(* IEC 61131-3 sources: deprecated-refusr-repo/samples (part 3) *)

(* ---- 2-MUX_whoso-sours-stout.st ---- *)
(*
This code implements a shuffled multiplexer with 2 control bits.
The control bits are: Data[3], Data[2]
The input bits are: Data[5], Data[1], Data[6], Data[4]

The symbolic expression is:
(((~(~(D[3]) & ~(D[2])) | D[5]) & (~(D[3] & ~(D[2])) | D[1])) & (~(~(D[3]) & D[2]) | D[6])) & (~(D[3] & D[2]) | D[4])

*)

FUNCTION_BLOCK F_CollectInput
  VAR_IN_OUT
      Data : ARRAY[1..10] OF BOOL;
  END_VAR
  VAR_INPUT
      TICK  : BOOL := 0;
      IN1   : BOOL := 0;
      IN2   : BOOL := 0;
      IN3   : BOOL := 0;
      IN4   : BOOL := 0;
      IN5   : BOOL := 0;
      RESET : BOOL := FALSE;
  END_VAR
  VAR_OUTPUT
      Finished : BOOL;
  END_VAR
  VAR
      j    : USINT := 1;
      tock : BOOL  := 0;
  END_VAR
  IF NOT RESET AND tock = NOT TICK THEN
      Data[j]   := IN1;
      Data[j+1] := IN2;
      Data[j+2] := IN3;
      Data[j+3] := IN4;
      Data[j+4] := IN5;
      j := j + 5;
      tock := TICK;
  ELSE
      j := 1;
      tock := 0;
  END_IF;
  Finished := (j > 10);
END_FUNCTION_BLOCK

PROGRAM Boiler
  VAR
    Data  : ARRAY[1..10] OF BOOL;
    Ready : BOOL;
    CollectInput : F_CollectInput;
  END_VAR
  VAR
    TICK     AT %IX1.0 : BOOL;
    IN1      AT %IX0.3 : BOOL;
    IN2      AT %IX0.4 : BOOL;
    IN3      AT %IX0.5 : BOOL;
    IN4      AT %IX0.6 : BOOL;
    IN5      AT %IX0.7 : BOOL;
    OutReady AT %QX0.0 : BOOL := FALSE;
    FeedNext AT %QX0.1 : BOOL := FALSE;
    Out      AT %QX0.2 : BOOL;
  END_VAR
  CollectInput(TICK:=TICK, IN1:=IN1, IN2:=IN2, IN3:=IN3, IN4:=IN4, IN5:=IN5);
  Ready := CollectInput.Finished;
  FeedNext := 1;
  IF Ready THEN
    Out := (((((NOT ((NOT D[3]) AND (NOT D[2]))) OR D[5]) AND ((NOT (D[3] AND (NOT D[2]))) OR D[1])) AND ((NOT ((NOT D[3]) AND D[2])) OR D[6])) AND ((NOT (D[3] AND D[2])) OR D[4]));
    OutReady := 1;
    CollectInput(RESET:=TRUE);
  END_IF;
END_PROGRAM

CONFIGURATION Config0
  RESOURCE Res0 ON PLC
    TASK task0(INTERVAL := T#20ms,PRIORITY := 0);
    PROGRAM instance0 WITH task0 : Boiler;
  END_RESOURCE
END_CONFIGURATION

(* ---- 2-MUX_wimpy-lubra-dopes.st ---- *)
(*
This code implements a shuffled multiplexer with 2 control bits.
The control bits are: Data[1], Data[5]
The input bits are: Data[3], Data[2], Data[4], Data[6]

The symbolic expression is:
(((~(~(D[1]) & ~(D[5])) | D[3]) & (~(D[1] & ~(D[5])) | D[2])) & (~(~(D[1]) & D[5]) | D[4])) & (~(D[1] & D[5]) | D[6])

*)

FUNCTION_BLOCK F_CollectInput
  VAR_IN_OUT
      Data : ARRAY[1..10] OF BOOL;
  END_VAR
  VAR_INPUT
      TICK  : BOOL := 0;
      IN1   : BOOL := 0;
      IN2   : BOOL := 0;
      IN3   : BOOL := 0;
      IN4   : BOOL := 0;
      IN5   : BOOL := 0;
      RESET : BOOL := FALSE;
  END_VAR
  VAR_OUTPUT
      Finished : BOOL;
  END_VAR
  VAR
      j    : USINT := 1;
      tock : BOOL  := 0;
  END_VAR
  IF NOT RESET AND tock = NOT TICK THEN
      Data[j]   := IN1;
      Data[j+1] := IN2;
      Data[j+2] := IN3;
      Data[j+3] := IN4;
      Data[j+4] := IN5;
      j := j + 5;
      tock := TICK;
  ELSE
      j := 1;
      tock := 0;
  END_IF;
  Finished := (j > 10);
END_FUNCTION_BLOCK

PROGRAM Boiler
  VAR
    Data  : ARRAY[1..10] OF BOOL;
    Ready : BOOL;
    CollectInput : F_CollectInput;
  END_VAR
  VAR
    TICK     AT %IX1.0 : BOOL;
    IN1      AT %IX0.3 : BOOL;
    IN2      AT %IX0.4 : BOOL;
    IN3      AT %IX0.5 : BOOL;
    IN4      AT %IX0.6 : BOOL;
    IN5      AT %IX0.7 : BOOL;
    OutReady AT %QX0.0 : BOOL := FALSE;
    FeedNext AT %QX0.1 : BOOL := FALSE;
    Out      AT %QX0.2 : BOOL;
  END_VAR
  CollectInput(TICK:=TICK, IN1:=IN1, IN2:=IN2, IN3:=IN3, IN4:=IN4, IN5:=IN5);
  Ready := CollectInput.Finished;
  FeedNext := 1;
  IF Ready THEN
    Out := (((((NOT ((NOT D[1]) AND (NOT D[5]))) OR D[3]) AND ((NOT (D[1] AND (NOT D[5]))) OR D[2])) AND ((NOT ((NOT D[1]) AND D[5])) OR D[4])) AND ((NOT (D[1] AND D[5])) OR D[6]));
    OutReady := 1;
    CollectInput(RESET:=TRUE);
  END_IF;
END_PROGRAM

CONFIGURATION Config0
  RESOURCE Res0 ON PLC
    TASK task0(INTERVAL := T#20ms,PRIORITY := 0);
    PROGRAM instance0 WITH task0 : Boiler;
  END_RESOURCE
END_CONFIGURATION

(* ---- 2-MUX_wolds-gists-resay.st ---- *)
(*
This code implements a shuffled multiplexer with 2 control bits.
The control bits are: Data[4], Data[2]
The input bits are: Data[5], Data[1], Data[3], Data[6]

The symbolic expression is:
(((~(~(D[4]) & ~(D[2])) | D[5]) & (~(D[4] & ~(D[2])) | D[1])) & (~(~(D[4]) & D[2]) | D[3])) & (~(D[4] & D[2]) | D[6])

*)

FUNCTION_BLOCK F_CollectInput
  VAR_IN_OUT
      Data : ARRAY[1..10] OF BOOL;
  END_VAR
  VAR_INPUT
      TICK  : BOOL := 0;
      IN1   : BOOL := 0;
      IN2   : BOOL := 0;
      IN3   : BOOL := 0;
      IN4   : BOOL := 0;
      IN5   : BOOL := 0;
      RESET : BOOL := FALSE;
  END_VAR
  VAR_OUTPUT
      Finished : BOOL;
  END_VAR
  VAR
      j    : USINT := 1;
      tock : BOOL  := 0;
  END_VAR
  IF NOT RESET AND tock = NOT TICK THEN
      Data[j]   := IN1;
      Data[j+1] := IN2;
      Data[j+2] := IN3;
      Data[j+3] := IN4;
      Data[j+4] := IN5;
      j := j + 5;
      tock := TICK;
  ELSE
      j := 1;
      tock := 0;
  END_IF;
  Finished := (j > 10);
END_FUNCTION_BLOCK

PROGRAM Boiler
  VAR
    Data  : ARRAY[1..10] OF BOOL;
    Ready : BOOL;
    CollectInput : F_CollectInput;
  END_VAR
  VAR
    TICK     AT %IX1.0 : BOOL;
    IN1      AT %IX0.3 : BOOL;
    IN2      AT %IX0.4 : BOOL;
    IN3      AT %IX0.5 : BOOL;
    IN4      AT %IX0.6 : BOOL;
    IN5      AT %IX0.7 : BOOL;
    OutReady AT %QX0.0 : BOOL := FALSE;
    FeedNext AT %QX0.1 : BOOL := FALSE;
    Out      AT %QX0.2 : BOOL;
  END_VAR
  CollectInput(TICK:=TICK, IN1:=IN1, IN2:=IN2, IN3:=IN3, IN4:=IN4, IN5:=IN5);
  Ready := CollectInput.Finished;
  FeedNext := 1;
  IF Ready THEN
    Out := (((((NOT ((NOT D[4]) AND (NOT D[2]))) OR D[5]) AND ((NOT (D[4] AND (NOT D[2]))) OR D[1])) AND ((NOT ((NOT D[4]) AND D[2])) OR D[3])) AND ((NOT (D[4] AND D[2])) OR D[6]));
    OutReady := 1;
    CollectInput(RESET:=TRUE);
  END_IF;
END_PROGRAM

CONFIGURATION Config0
  RESOURCE Res0 ON PLC
    TASK task0(INTERVAL := T#20ms,PRIORITY := 0);
    PROGRAM instance0 WITH task0 : Boiler;
  END_RESOURCE
END_CONFIGURATION

(* ---- 2-MUX_yella-trams-woken.st ---- *)
(*
This code implements a shuffled multiplexer with 2 control bits.
The control bits are: Data[1], Data[2]
The input bits are: Data[3], Data[5], Data[6], Data[4]

The symbolic expression is:
(((~(~(D[1]) & ~(D[2])) | D[3]) & (~(D[1] & ~(D[2])) | D[5])) & (~(~(D[1]) & D[2]) | D[6])) & (~(D[1] & D[2]) | D[4])

*)

FUNCTION_BLOCK F_CollectInput
  VAR_IN_OUT
      Data : ARRAY[1..10] OF BOOL;
  END_VAR
  VAR_INPUT
      TICK  : BOOL := 0;
      IN1   : BOOL := 0;
      IN2   : BOOL := 0;
      IN3   : BOOL := 0;
      IN4   : BOOL := 0;
      IN5   : BOOL := 0;
      RESET : BOOL := FALSE;
  END_VAR
  VAR_OUTPUT
      Finished : BOOL;
  END_VAR
  VAR
      j    : USINT := 1;
      tock : BOOL  := 0;
  END_VAR
  IF NOT RESET AND tock = NOT TICK THEN
      Data[j]   := IN1;
      Data[j+1] := IN2;
      Data[j+2] := IN3;
      Data[j+3] := IN4;
      Data[j+4] := IN5;
      j := j + 5;
      tock := TICK;
  ELSE
      j := 1;
      tock := 0;
  END_IF;
  Finished := (j > 10);
END_FUNCTION_BLOCK

PROGRAM Boiler
  VAR
    Data  : ARRAY[1..10] OF BOOL;
    Ready : BOOL;
    CollectInput : F_CollectInput;
  END_VAR
  VAR
    TICK     AT %IX1.0 : BOOL;
    IN1      AT %IX0.3 : BOOL;
    IN2      AT %IX0.4 : BOOL;
    IN3      AT %IX0.5 : BOOL;
    IN4      AT %IX0.6 : BOOL;
    IN5      AT %IX0.7 : BOOL;
    OutReady AT %QX0.0 : BOOL := FALSE;
    FeedNext AT %QX0.1 : BOOL := FALSE;
    Out      AT %QX0.2 : BOOL;
  END_VAR
  CollectInput(TICK:=TICK, IN1:=IN1, IN2:=IN2, IN3:=IN3, IN4:=IN4, IN5:=IN5);
  Ready := CollectInput.Finished;
  FeedNext := 1;
  IF Ready THEN
    Out := (((((NOT ((NOT D[1]) AND (NOT D[2]))) OR D[3]) AND ((NOT (D[1] AND (NOT D[2]))) OR D[5])) AND ((NOT ((NOT D[1]) AND D[2])) OR D[6])) AND ((NOT (D[1] AND D[2])) OR D[4]));
    OutReady := 1;
    CollectInput(RESET:=TRUE);
  END_IF;
END_PROGRAM

CONFIGURATION Config0
  RESOURCE Res0 ON PLC
    TASK task0(INTERVAL := T#20ms,PRIORITY := 0);
    PROGRAM instance0 WITH task0 : Boiler;
  END_RESOURCE
END_CONFIGURATION

(* ---- 2-MUX_yoyos-blast-cameo.st ---- *)
(*
This code implements a shuffled multiplexer with 2 control bits.
The control bits are: Data[3], Data[2]
The input bits are: Data[1], Data[4], Data[5], Data[6]

The symbolic expression is:
(((~(~(D[3]) & ~(D[2])) | D[1]) & (~(D[3] & ~(D[2])) | D[4])) & (~(~(D[3]) & D[2]) | D[5])) & (~(D[3] & D[2]) | D[6])

*)

FUNCTION_BLOCK F_CollectInput
  VAR_IN_OUT
      Data : ARRAY[1..10] OF BOOL;
  END_VAR
  VAR_INPUT
      TICK  : BOOL := 0;
      IN1   : BOOL := 0;
      IN2   : BOOL := 0;
      IN3   : BOOL := 0;
      IN4   : BOOL := 0;
      IN5   : BOOL := 0;
      RESET : BOOL := FALSE;
  END_VAR
  VAR_OUTPUT
      Finished : BOOL;
  END_VAR
  VAR
      j    : USINT := 1;
      tock : BOOL  := 0;
  END_VAR
  IF NOT RESET AND tock = NOT TICK THEN
      Data[j]   := IN1;
      Data[j+1] := IN2;
      Data[j+2] := IN3;
      Data[j+3] := IN4;
      Data[j+4] := IN5;
      j := j + 5;
      tock := TICK;
  ELSE
      j := 1;
      tock := 0;
  END_IF;
  Finished := (j > 10);
END_FUNCTION_BLOCK

PROGRAM Boiler
  VAR
    Data  : ARRAY[1..10] OF BOOL;
    Ready : BOOL;
    CollectInput : F_CollectInput;
  END_VAR
  VAR
    TICK     AT %IX1.0 : BOOL;
    IN1      AT %IX0.3 : BOOL;
    IN2      AT %IX0.4 : BOOL;
    IN3      AT %IX0.5 : BOOL;
    IN4      AT %IX0.6 : BOOL;
    IN5      AT %IX0.7 : BOOL;
    OutReady AT %QX0.0 : BOOL := FALSE;
    FeedNext AT %QX0.1 : BOOL := FALSE;
    Out      AT %QX0.2 : BOOL;
  END_VAR
  CollectInput(TICK:=TICK, IN1:=IN1, IN2:=IN2, IN3:=IN3, IN4:=IN4, IN5:=IN5);
  Ready := CollectInput.Finished;
  FeedNext := 1;
  IF Ready THEN
    Out := (((((NOT ((NOT D[3]) AND (NOT D[2]))) OR D[1]) AND ((NOT (D[3] AND (NOT D[2]))) OR D[4])) AND ((NOT ((NOT D[3]) AND D[2])) OR D[5])) AND ((NOT (D[3] AND D[2])) OR D[6]));
    OutReady := 1;
    CollectInput(RESET:=TRUE);
  END_IF;
END_PROGRAM

CONFIGURATION Config0
  RESOURCE Res0 ON PLC
    TASK task0(INTERVAL := T#20ms,PRIORITY := 0);
    PROGRAM instance0 WITH task0 : Boiler;
  END_RESOURCE
END_CONFIGURATION

(* ---- 2-MUX_yurts-tippy-sayer.st ---- *)
(*
This code implements a shuffled multiplexer with 2 control bits.
The control bits are: Data[3], Data[1]
The input bits are: Data[4], Data[2], Data[5], Data[6]

The symbolic expression is:
(((~(~(D[3]) & ~(D[1])) | D[4]) & (~(D[3] & ~(D[1])) | D[2])) & (~(~(D[3]) & D[1]) | D[5])) & (~(D[3] & D[1]) | D[6])

*)

FUNCTION_BLOCK F_CollectInput
  VAR_IN_OUT
      Data : ARRAY[1..10] OF BOOL;
  END_VAR
  VAR_INPUT
      TICK  : BOOL := 0;
      IN1   : BOOL := 0;
      IN2   : BOOL := 0;
      IN3   : BOOL := 0;
      IN4   : BOOL := 0;
      IN5   : BOOL := 0;
      RESET : BOOL := FALSE;
  END_VAR
  VAR_OUTPUT
      Finished : BOOL;
  END_VAR
  VAR
      j    : USINT := 1;
      tock : BOOL  := 0;
  END_VAR
  IF NOT RESET AND tock = NOT TICK THEN
      Data[j]   := IN1;
      Data[j+1] := IN2;
      Data[j+2] := IN3;
      Data[j+3] := IN4;
      Data[j+4] := IN5;
      j := j + 5;
      tock := TICK;
  ELSE
      j := 1;
      tock := 0;
  END_IF;
  Finished := (j > 10);
END_FUNCTION_BLOCK

PROGRAM Boiler
  VAR
    Data  : ARRAY[1..10] OF BOOL;
    Ready : BOOL;
    CollectInput : F_CollectInput;
  END_VAR
  VAR
    TICK     AT %IX1.0 : BOOL;
    IN1      AT %IX0.3 : BOOL;
    IN2      AT %IX0.4 : BOOL;
    IN3      AT %IX0.5 : BOOL;
    IN4      AT %IX0.6 : BOOL;
    IN5      AT %IX0.7 : BOOL;
    OutReady AT %QX0.0 : BOOL := FALSE;
    FeedNext AT %QX0.1 : BOOL := FALSE;
    Out      AT %QX0.2 : BOOL;
  END_VAR
  CollectInput(TICK:=TICK, IN1:=IN1, IN2:=IN2, IN3:=IN3, IN4:=IN4, IN5:=IN5);
  Ready := CollectInput.Finished;
  FeedNext := 1;
  IF Ready THEN
    Out := (((((NOT ((NOT D[3]) AND (NOT D[1]))) OR D[4]) AND ((NOT (D[3] AND (NOT D[1]))) OR D[2])) AND ((NOT ((NOT D[3]) AND D[1])) OR D[5])) AND ((NOT (D[3] AND D[1])) OR D[6]));
    OutReady := 1;
    CollectInput(RESET:=TRUE);
  END_IF;
END_PROGRAM

CONFIGURATION Config0
  RESOURCE Res0 ON PLC
    TASK task0(INTERVAL := T#20ms,PRIORITY := 0);
    PROGRAM instance0 WITH task0 : Boiler;
  END_RESOURCE
END_CONFIGURATION

(* ---- 2-MUX_zebus-trove-teals.st ---- *)
(*
This code implements a shuffled multiplexer with 2 control bits.
The control bits are: Data[2], Data[1]
The input bits are: Data[5], Data[6], Data[3], Data[4]

The symbolic expression is:
(((~(~(D[2]) & ~(D[1])) | D[5]) & (~(D[2] & ~(D[1])) | D[6])) & (~(~(D[2]) & D[1]) | D[3])) & (~(D[2] & D[1]) | D[4])

*)

FUNCTION_BLOCK F_CollectInput
  VAR_IN_OUT
      Data : ARRAY[1..10] OF BOOL;
  END_VAR
  VAR_INPUT
      TICK  : BOOL := 0;
      IN1   : BOOL := 0;
      IN2   : BOOL := 0;
      IN3   : BOOL := 0;
      IN4   : BOOL := 0;
      IN5   : BOOL := 0;
      RESET : BOOL := FALSE;
  END_VAR
  VAR_OUTPUT
      Finished : BOOL;
  END_VAR
  VAR
      j    : USINT := 1;
      tock : BOOL  := 0;
  END_VAR
  IF NOT RESET AND tock = NOT TICK THEN
      Data[j]   := IN1;
      Data[j+1] := IN2;
      Data[j+2] := IN3;
      Data[j+3] := IN4;
      Data[j+4] := IN5;
      j := j + 5;
      tock := TICK;
  ELSE
      j := 1;
      tock := 0;
  END_IF;
  Finished := (j > 10);
END_FUNCTION_BLOCK

PROGRAM Boiler
  VAR
    Data  : ARRAY[1..10] OF BOOL;
    Ready : BOOL;
    CollectInput : F_CollectInput;
  END_VAR
  VAR
    TICK     AT %IX1.0 : BOOL;
    IN1      AT %IX0.3 : BOOL;
    IN2      AT %IX0.4 : BOOL;
    IN3      AT %IX0.5 : BOOL;
    IN4      AT %IX0.6 : BOOL;
    IN5      AT %IX0.7 : BOOL;
    OutReady AT %QX0.0 : BOOL := FALSE;
    FeedNext AT %QX0.1 : BOOL := FALSE;
    Out      AT %QX0.2 : BOOL;
  END_VAR
  CollectInput(TICK:=TICK, IN1:=IN1, IN2:=IN2, IN3:=IN3, IN4:=IN4, IN5:=IN5);
  Ready := CollectInput.Finished;
  FeedNext := 1;
  IF Ready THEN
    Out := (((((NOT ((NOT D[2]) AND (NOT D[1]))) OR D[5]) AND ((NOT (D[2] AND (NOT D[1]))) OR D[6])) AND ((NOT ((NOT D[2]) AND D[1])) OR D[3])) AND ((NOT (D[2] AND D[1])) OR D[4]));
    OutReady := 1;
    CollectInput(RESET:=TRUE);
  END_IF;
END_PROGRAM

CONFIGURATION Config0
  RESOURCE Res0 ON PLC
    TASK task0(INTERVAL := T#20ms,PRIORITY := 0);
    PROGRAM instance0 WITH task0 : Boiler;
  END_RESOURCE
END_CONFIGURATION

(* ---- 2-MUX_zebus-whiny-fares.st ---- *)
(*
This code implements a shuffled multiplexer with 2 control bits.
The control bits are: Data[1], Data[2]
The input bits are: Data[3], Data[4], Data[5], Data[6]

The symbolic expression is:
(((~(~(D[1]) & ~(D[2])) | D[3]) & (~(D[1] & ~(D[2])) | D[4])) & (~(~(D[1]) & D[2]) | D[5])) & (~(D[1] & D[2]) | D[6])

*)

FUNCTION_BLOCK F_CollectInput
  VAR_IN_OUT
      Data : ARRAY[1..10] OF BOOL;
  END_VAR
  VAR_INPUT
      TICK  : BOOL := 0;
      IN1   : BOOL := 0;
      IN2   : BOOL := 0;
      IN3   : BOOL := 0;
      IN4   : BOOL := 0;
      IN5   : BOOL := 0;
      RESET : BOOL := FALSE;
  END_VAR
  VAR_OUTPUT
      Finished : BOOL;
  END_VAR
  VAR
      j    : USINT := 1;
      tock : BOOL  := 0;
  END_VAR
  IF NOT RESET AND tock = NOT TICK THEN
      Data[j]   := IN1;
      Data[j+1] := IN2;
      Data[j+2] := IN3;
      Data[j+3] := IN4;
      Data[j+4] := IN5;
      j := j + 5;
      tock := TICK;
  ELSE
      j := 1;
      tock := 0;
  END_IF;
  Finished := (j > 10);
END_FUNCTION_BLOCK

PROGRAM Boiler
  VAR
    Data  : ARRAY[1..10] OF BOOL;
    Ready : BOOL;
    CollectInput : F_CollectInput;
  END_VAR
  VAR
    TICK     AT %IX1.0 : BOOL;
    IN1      AT %IX0.3 : BOOL;
    IN2      AT %IX0.4 : BOOL;
    IN3      AT %IX0.5 : BOOL;
    IN4      AT %IX0.6 : BOOL;
    IN5      AT %IX0.7 : BOOL;
    OutReady AT %QX0.0 : BOOL := FALSE;
    FeedNext AT %QX0.1 : BOOL := FALSE;
    Out      AT %QX0.2 : BOOL;
  END_VAR
  CollectInput(TICK:=TICK, IN1:=IN1, IN2:=IN2, IN3:=IN3, IN4:=IN4, IN5:=IN5);
  Ready := CollectInput.Finished;
  FeedNext := 1;
  IF Ready THEN
    Out := (((((NOT ((NOT D[1]) AND (NOT D[2]))) OR D[3]) AND ((NOT (D[1] AND (NOT D[2]))) OR D[4])) AND ((NOT ((NOT D[1]) AND D[2])) OR D[5])) AND ((NOT (D[1] AND D[2])) OR D[6]));
    OutReady := 1;
    CollectInput(RESET:=TRUE);
  END_IF;
END_PROGRAM

CONFIGURATION Config0
  RESOURCE Res0 ON PLC
    TASK task0(INTERVAL := T#20ms,PRIORITY := 0);
    PROGRAM instance0 WITH task0 : Boiler;
  END_RESOURCE
END_CONFIGURATION

(* ---- 3-MUX_acked-palls-seven.st ---- *)
(*
This code implements a shuffled multiplexer with 3 control bits.
The control bits are: Data[2], Data[1], Data[3]
The input bits are: Data[4], Data[6], Data[7], Data[5], Data[8], Data[9], Data[11], Data[10]

The symbolic expression is:
(((((((~((~(D[2]) & ~(D[1])) & ~(D[3])) | D[4]) & (~((D[2] & ~(D[1])) & ~(D[3])) | D[6])) & (~((~(D[2]) & D[1]) & ~(D[3])) | D[7])) & (~((D[2] & D[1]) & ~(D[3])) | D[5])) & (~((~(D[2]) & ~(D[1])) & D[3]) | D[8])) & (~((D[2] & ~(D[1])) & D[3]) | D[9])) & (~((~(D[2]) & D[1]) & D[3]) | D[11])) & (~((D[2] & D[1]) & D[3]) | D[10])

*)

FUNCTION_BLOCK F_CollectInput
  VAR_IN_OUT
      Data : ARRAY[1..15] OF BOOL;
  END_VAR
  VAR_INPUT
      TICK  : BOOL := 0;
      IN1   : BOOL := 0;
      IN2   : BOOL := 0;
      IN3   : BOOL := 0;
      IN4   : BOOL := 0;
      IN5   : BOOL := 0;
      RESET : BOOL := FALSE;
  END_VAR
  VAR_OUTPUT
      Finished : BOOL;
  END_VAR
  VAR
      j    : USINT := 1;
      tock : BOOL  := 0;
  END_VAR
  IF NOT RESET AND tock = NOT TICK THEN
      Data[j]   := IN1;
      Data[j+1] := IN2;
      Data[j+2] := IN3;
      Data[j+3] := IN4;
      Data[j+4] := IN5;
      j := j + 5;
      tock := TICK;
  ELSE
      j := 1;
      tock := 0;
  END_IF;
  Finished := (j > 15);
END_FUNCTION_BLOCK

PROGRAM Boiler
  VAR
    Data  : ARRAY[1..15] OF BOOL;
    Ready : BOOL;
    CollectInput : F_CollectInput;
  END_VAR
  VAR
    TICK     AT %IX1.0 : BOOL;
    IN1      AT %IX0.3 : BOOL;
    IN2      AT %IX0.4 : BOOL;
    IN3      AT %IX0.5 : BOOL;
    IN4      AT %IX0.6 : BOOL;
    IN5      AT %IX0.7 : BOOL;
    OutReady AT %QX0.0 : BOOL := FALSE;
    FeedNext AT %QX0.1 : BOOL := FALSE;
    Out      AT %QX0.2 : BOOL;
  END_VAR
  CollectInput(TICK:=TICK, IN1:=IN1, IN2:=IN2, IN3:=IN3, IN4:=IN4, IN5:=IN5);
  Ready := CollectInput.Finished;
  FeedNext := 1;
  IF Ready THEN
    Out := (((((((((NOT (((NOT D[2]) AND (NOT D[1])) AND (NOT D[3]))) OR D[4]) AND ((NOT ((D[2] AND (NOT D[1])) AND (NOT D[3]))) OR D[6])) AND ((NOT (((NOT D[2]) AND D[1]) AND (NOT D[3]))) OR D[7])) AND ((NOT ((D[2] AND D[1]) AND (NOT D[3]))) OR D[5])) AND ((NOT (((NOT D[2]) AND (NOT D[1])) AND D[3])) OR D[8])) AND ((NOT ((D[2] AND (NOT D[1])) AND D[3])) OR D[9])) AND ((NOT (((NOT D[2]) AND D[1]) AND D[3])) OR D[11])) AND ((NOT ((D[2] AND D[1]) AND D[3])) OR D[10]));
    OutReady := 1;
    CollectInput(RESET:=TRUE);
  END_IF;
END_PROGRAM

CONFIGURATION Config0
  RESOURCE Res0 ON PLC
    TASK task0(INTERVAL := T#20ms,PRIORITY := 0);
    PROGRAM instance0 WITH task0 : Boiler;
  END_RESOURCE
END_CONFIGURATION

(* ---- 3-MUX_alums-tends-demon.st ---- *)
(*
This code implements a shuffled multiplexer with 3 control bits.
The control bits are: Data[1], Data[3], Data[6]
The input bits are: Data[4], Data[9], Data[5], Data[2], Data[7], Data[8], Data[10], Data[11]

The symbolic expression is:
(((((((~((~(D[1]) & ~(D[3])) & ~(D[6])) | D[4]) & (~((D[1] & ~(D[3])) & ~(D[6])) | D[9])) & (~((~(D[1]) & D[3]) & ~(D[6])) | D[5])) & (~((D[1] & D[3]) & ~(D[6])) | D[2])) & (~((~(D[1]) & ~(D[3])) & D[6]) | D[7])) & (~((D[1] & ~(D[3])) & D[6]) | D[8])) & (~((~(D[1]) & D[3]) & D[6]) | D[10])) & (~((D[1] & D[3]) & D[6]) | D[11])

*)

FUNCTION_BLOCK F_CollectInput
  VAR_IN_OUT
      Data : ARRAY[1..15] OF BOOL;
  END_VAR
  VAR_INPUT
      TICK  : BOOL := 0;
      IN1   : BOOL := 0;
      IN2   : BOOL := 0;
      IN3   : BOOL := 0;
      IN4   : BOOL := 0;
      IN5   : BOOL := 0;
      RESET : BOOL := FALSE;
  END_VAR
  VAR_OUTPUT
      Finished : BOOL;
  END_VAR
  VAR
      j    : USINT := 1;
      tock : BOOL  := 0;
  END_VAR
  IF NOT RESET AND tock = NOT TICK THEN
      Data[j]   := IN1;
      Data[j+1] := IN2;
      Data[j+2] := IN3;
      Data[j+3] := IN4;
      Data[j+4] := IN5;
      j := j + 5;
      tock := TICK;
  ELSE
      j := 1;
      tock := 0;
  END_IF;
  Finished := (j > 15);
END_FUNCTION_BLOCK

PROGRAM Boiler
  VAR
    Data  : ARRAY[1..15] OF BOOL;
    Ready : BOOL;
    CollectInput : F_CollectInput;
  END_VAR
  VAR
    TICK     AT %IX1.0 : BOOL;
    IN1      AT %IX0.3 : BOOL;
    IN2      AT %IX0.4 : BOOL;
    IN3      AT %IX0.5 : BOOL;
    IN4      AT %IX0.6 : BOOL;
    IN5      AT %IX0.7 : BOOL;
    OutReady AT %QX0.0 : BOOL := FALSE;
    FeedNext AT %QX0.1 : BOOL := FALSE;
    Out      AT %QX0.2 : BOOL;
  END_VAR
  CollectInput(TICK:=TICK, IN1:=IN1, IN2:=IN2, IN3:=IN3, IN4:=IN4, IN5:=IN5);
  Ready := CollectInput.Finished;
  FeedNext := 1;
  IF Ready THEN
    Out := (((((((((NOT (((NOT D[1]) AND (NOT D[3])) AND (NOT D[6]))) OR D[4]) AND ((NOT ((D[1] AND (NOT D[3])) AND (NOT D[6]))) OR D[9])) AND ((NOT (((NOT D[1]) AND D[3]) AND (NOT D[6]))) OR D[5])) AND ((NOT ((D[1] AND D[3]) AND (NOT D[6]))) OR D[2])) AND ((NOT (((NOT D[1]) AND (NOT D[3])) AND D[6])) OR D[7])) AND ((NOT ((D[1] AND (NOT D[3])) AND D[6])) OR D[8])) AND ((NOT (((NOT D[1]) AND D[3]) AND D[6])) OR D[10])) AND ((NOT ((D[1] AND D[3]) AND D[6])) OR D[11]));
    OutReady := 1;
    CollectInput(RESET:=TRUE);
  END_IF;
END_PROGRAM

CONFIGURATION Config0
  RESOURCE Res0 ON PLC
    TASK task0(INTERVAL := T#20ms,PRIORITY := 0);
    PROGRAM instance0 WITH task0 : Boiler;
  END_RESOURCE
END_CONFIGURATION

(* ---- 3-MUX_annex-saucy-first.st ---- *)
(*
This code implements a shuffled multiplexer with 3 control bits.
The control bits are: Data[2], Data[1], Data[5]
The input bits are: Data[3], Data[6], Data[4], Data[7], Data[8], Data[9], Data[10], Data[11]

The symbolic expression is:
(((((((~((~(D[2]) & ~(D[1])) & ~(D[5])) | D[3]) & (~((D[2] & ~(D[1])) & ~(D[5])) | D[6])) & (~((~(D[2]) & D[1]) & ~(D[5])) | D[4])) & (~((D[2] & D[1]) & ~(D[5])) | D[7])) & (~((~(D[2]) & ~(D[1])) & D[5]) | D[8])) & (~((D[2] & ~(D[1])) & D[5]) | D[9])) & (~((~(D[2]) & D[1]) & D[5]) | D[10])) & (~((D[2] & D[1]) & D[5]) | D[11])

*)

FUNCTION_BLOCK F_CollectInput
  VAR_IN_OUT
      Data : ARRAY[1..15] OF BOOL;
  END_VAR
  VAR_INPUT
      TICK  : BOOL := 0;
      IN1   : BOOL := 0;
      IN2   : BOOL := 0;
      IN3   : BOOL := 0;
      IN4   : BOOL := 0;
      IN5   : BOOL := 0;
      RESET : BOOL := FALSE;
  END_VAR
  VAR_OUTPUT
      Finished : BOOL;
  END_VAR
  VAR
      j    : USINT := 1;
      tock : BOOL  := 0;
  END_VAR
  IF NOT RESET AND tock = NOT TICK THEN
      Data[j]   := IN1;
      Data[j+1] := IN2;
      Data[j+2] := IN3;
      Data[j+3] := IN4;
      Data[j+4] := IN5;
      j := j + 5;
      tock := TICK;
  ELSE
      j := 1;
      tock := 0;
  END_IF;
  Finished := (j > 15);
END_FUNCTION_BLOCK

PROGRAM Boiler
  VAR
    Data  : ARRAY[1..15] OF BOOL;
    Ready : BOOL;
    CollectInput : F_CollectInput;
  END_VAR
  VAR
    TICK     AT %IX1.0 : BOOL;
    IN1      AT %IX0.3 : BOOL;
    IN2      AT %IX0.4 : BOOL;
    IN3      AT %IX0.5 : BOOL;
    IN4      AT %IX0.6 : BOOL;
    IN5      AT %IX0.7 : BOOL;
    OutReady AT %QX0.0 : BOOL := FALSE;
    FeedNext AT %QX0.1 : BOOL := FALSE;
    Out      AT %QX0.2 : BOOL;
  END_VAR
  CollectInput(TICK:=TICK, IN1:=IN1, IN2:=IN2, IN3:=IN3, IN4:=IN4, IN5:=IN5);
  Ready := CollectInput.Finished;
  FeedNext := 1;
  IF Ready THEN
    Out := (((((((((NOT (((NOT D[2]) AND (NOT D[1])) AND (NOT D[5]))) OR D[3]) AND ((NOT ((D[2] AND (NOT D[1])) AND (NOT D[5]))) OR D[6])) AND ((NOT (((NOT D[2]) AND D[1]) AND (NOT D[5]))) OR D[4])) AND ((NOT ((D[2] AND D[1]) AND (NOT D[5]))) OR D[7])) AND ((NOT (((NOT D[2]) AND (NOT D[1])) AND D[5])) OR D[8])) AND ((NOT ((D[2] AND (NOT D[1])) AND D[5])) OR D[9])) AND ((NOT (((NOT D[2]) AND D[1]) AND D[5])) OR D[10])) AND ((NOT ((D[2] AND D[1]) AND D[5])) OR D[11]));
    OutReady := 1;
    CollectInput(RESET:=TRUE);
  END_IF;
END_PROGRAM

CONFIGURATION Config0
  RESOURCE Res0 ON PLC
    TASK task0(INTERVAL := T#20ms,PRIORITY := 0);
    PROGRAM instance0 WITH task0 : Boiler;
  END_RESOURCE
END_CONFIGURATION

(* ---- 3-MUX_antic-lucks-mould.st ---- *)
(*
This code implements a shuffled multiplexer with 3 control bits.
The control bits are: Data[2], Data[7], Data[1]
The input bits are: Data[3], Data[5], Data[6], Data[4], Data[8], Data[9], Data[10], Data[11]

The symbolic expression is:
(((((((~((~(D[2]) & ~(D[7])) & ~(D[1])) | D[3]) & (~((D[2] & ~(D[7])) & ~(D[1])) | D[5])) & (~((~(D[2]) & D[7]) & ~(D[1])) | D[6])) & (~((D[2] & D[7]) & ~(D[1])) | D[4])) & (~((~(D[2]) & ~(D[7])) & D[1]) | D[8])) & (~((D[2] & ~(D[7])) & D[1]) | D[9])) & (~((~(D[2]) & D[7]) & D[1]) | D[10])) & (~((D[2] & D[7]) & D[1]) | D[11])

*)

FUNCTION_BLOCK F_CollectInput
  VAR_IN_OUT
      Data : ARRAY[1..15] OF BOOL;
  END_VAR
  VAR_INPUT
      TICK  : BOOL := 0;
      IN1   : BOOL := 0;
      IN2   : BOOL := 0;
      IN3   : BOOL := 0;
      IN4   : BOOL := 0;
      IN5   : BOOL := 0;
      RESET : BOOL := FALSE;
  END_VAR
  VAR_OUTPUT
      Finished : BOOL;
  END_VAR
  VAR
      j    : USINT := 1;
      tock : BOOL  := 0;
  END_VAR
  IF NOT RESET AND tock = NOT TICK THEN
      Data[j]   := IN1;
      Data[j+1] := IN2;
      Data[j+2] := IN3;
      Data[j+3] := IN4;
      Data[j+4] := IN5;
      j := j + 5;
      tock := TICK;
  ELSE
      j := 1;
      tock := 0;
  END_IF;
  Finished := (j > 15);
END_FUNCTION_BLOCK

PROGRAM Boiler
  VAR
    Data  : ARRAY[1..15] OF BOOL;
    Ready : BOOL;
    CollectInput : F_CollectInput;
  END_VAR
  VAR
    TICK     AT %IX1.0 : BOOL;
    IN1      AT %IX0.3 : BOOL;
    IN2      AT %IX0.4 : BOOL;
    IN3      AT %IX0.5 : BOOL;
    IN4      AT %IX0.6 : BOOL;
    IN5      AT %IX0.7 : BOOL;
    OutReady AT %QX0.0 : BOOL := FALSE;
    FeedNext AT %QX0.1 : BOOL := FALSE;
    Out      AT %QX0.2 : BOOL;
  END_VAR
  CollectInput(TICK:=TICK, IN1:=IN1, IN2:=IN2, IN3:=IN3, IN4:=IN4, IN5:=IN5);
  Ready := CollectInput.Finished;
  FeedNext := 1;
  IF Ready THEN
    Out := (((((((((NOT (((NOT D[2]) AND (NOT D[7])) AND (NOT D[1]))) OR D[3]) AND ((NOT ((D[2] AND (NOT D[7])) AND (NOT D[1]))) OR D[5])) AND ((NOT (((NOT D[2]) AND D[7]) AND (NOT D[1]))) OR D[6])) AND ((NOT ((D[2] AND D[7]) AND (NOT D[1]))) OR D[4])) AND ((NOT (((NOT D[2]) AND (NOT D[7])) AND D[1])) OR D[8])) AND ((NOT ((D[2] AND (NOT D[7])) AND D[1])) OR D[9])) AND ((NOT (((NOT D[2]) AND D[7]) AND D[1])) OR D[10])) AND ((NOT ((D[2] AND D[7]) AND D[1])) OR D[11]));
    OutReady := 1;
    CollectInput(RESET:=TRUE);
  END_IF;
END_PROGRAM

CONFIGURATION Config0
  RESOURCE Res0 ON PLC
    TASK task0(INTERVAL := T#20ms,PRIORITY := 0);
    PROGRAM instance0 WITH task0 : Boiler;
  END_RESOURCE
END_CONFIGURATION

(* ---- 3-MUX_apian-braes-rolls.st ---- *)
(*
This code implements a shuffled multiplexer with 3 control bits.
The control bits are: Data[2], Data[3], Data[1]
The input bits are: Data[4], Data[6], Data[5], Data[7], Data[10], Data[8], Data[9], Data[11]

The symbolic expression is:
(((((((~((~(D[2]) & ~(D[3])) & ~(D[1])) | D[4]) & (~((D[2] & ~(D[3])) & ~(D[1])) | D[6])) & (~((~(D[2]) & D[3]) & ~(D[1])) | D[5])) & (~((D[2] & D[3]) & ~(D[1])) | D[7])) & (~((~(D[2]) & ~(D[3])) & D[1]) | D[10])) & (~((D[2] & ~(D[3])) & D[1]) | D[8])) & (~((~(D[2]) & D[3]) & D[1]) | D[9])) & (~((D[2] & D[3]) & D[1]) | D[11])

*)

FUNCTION_BLOCK F_CollectInput
  VAR_IN_OUT
      Data : ARRAY[1..15] OF BOOL;
  END_VAR
  VAR_INPUT
      TICK  : BOOL := 0;
      IN1   : BOOL := 0;
      IN2   : BOOL := 0;
      IN3   : BOOL := 0;
      IN4   : BOOL := 0;
      IN5   : BOOL := 0;
      RESET : BOOL := FALSE;
  END_VAR
  VAR_OUTPUT
      Finished : BOOL;
  END_VAR
  VAR
      j    : USINT := 1;
      tock : BOOL  := 0;
  END_VAR
  IF NOT RESET AND tock = NOT TICK THEN
      Data[j]   := IN1;
      Data[j+1] := IN2;
      Data[j+2] := IN3;
      Data[j+3] := IN4;
      Data[j+4] := IN5;
      j := j + 5;
      tock := TICK;
  ELSE
      j := 1;
      tock := 0;
  END_IF;
  Finished := (j > 15);
END_FUNCTION_BLOCK

PROGRAM Boiler
  VAR
    Data  : ARRAY[1..15] OF BOOL;
    Ready : BOOL;
    CollectInput : F_CollectInput;
  END_VAR
  VAR
    TICK     AT %IX1.0 : BOOL;
    IN1      AT %IX0.3 : BOOL;
    IN2      AT %IX0.4 : BOOL;
    IN3      AT %IX0.5 : BOOL;
    IN4      AT %IX0.6 : BOOL;
    IN5      AT %IX0.7 : BOOL;
    OutReady AT %QX0.0 : BOOL := FALSE;
    FeedNext AT %QX0.1 : BOOL := FALSE;
    Out      AT %QX0.2 : BOOL;
  END_VAR
  CollectInput(TICK:=TICK, IN1:=IN1, IN2:=IN2, IN3:=IN3, IN4:=IN4, IN5:=IN5);
  Ready := CollectInput.Finished;
  FeedNext := 1;
  IF Ready THEN
    Out := (((((((((NOT (((NOT D[2]) AND (NOT D[3])) AND (NOT D[1]))) OR D[4]) AND ((NOT ((D[2] AND (NOT D[3])) AND (NOT D[1]))) OR D[6])) AND ((NOT (((NOT D[2]) AND D[3]) AND (NOT D[1]))) OR D[5])) AND ((NOT ((D[2] AND D[3]) AND (NOT D[1]))) OR D[7])) AND ((NOT (((NOT D[2]) AND (NOT D[3])) AND D[1])) OR D[10])) AND ((NOT ((D[2] AND (NOT D[3])) AND D[1])) OR D[8])) AND ((NOT (((NOT D[2]) AND D[3]) AND D[1])) OR D[9])) AND ((NOT ((D[2] AND D[3]) AND D[1])) OR D[11]));
    OutReady := 1;
    CollectInput(RESET:=TRUE);
  END_IF;
END_PROGRAM

CONFIGURATION Config0
  RESOURCE Res0 ON PLC
    TASK task0(INTERVAL := T#20ms,PRIORITY := 0);
    PROGRAM instance0 WITH task0 : Boiler;
  END_RESOURCE
END_CONFIGURATION

(* ---- 3-MUX_aping-spark-squad.st ---- *)
(*
This code implements a shuffled multiplexer with 3 control bits.
The control bits are: Data[5], Data[2], Data[1]
The input bits are: Data[4], Data[3], Data[6], Data[7], Data[8], Data[10], Data[9], Data[11]

The symbolic expression is:
(((((((~((~(D[5]) & ~(D[2])) & ~(D[1])) | D[4]) & (~((D[5] & ~(D[2])) & ~(D[1])) | D[3])) & (~((~(D[5]) & D[2]) & ~(D[1])) | D[6])) & (~((D[5] & D[2]) & ~(D[1])) | D[7])) & (~((~(D[5]) & ~(D[2])) & D[1]) | D[8])) & (~((D[5] & ~(D[2])) & D[1]) | D[10])) & (~((~(D[5]) & D[2]) & D[1]) | D[9])) & (~((D[5] & D[2]) & D[1]) | D[11])

*)

FUNCTION_BLOCK F_CollectInput
  VAR_IN_OUT
      Data : ARRAY[1..15] OF BOOL;
  END_VAR
  VAR_INPUT
      TICK  : BOOL := 0;
      IN1   : BOOL := 0;
      IN2   : BOOL := 0;
      IN3   : BOOL := 0;
      IN4   : BOOL := 0;
      IN5   : BOOL := 0;
      RESET : BOOL := FALSE;
  END_VAR
  VAR_OUTPUT
      Finished : BOOL;
  END_VAR
  VAR
      j    : USINT := 1;
      tock : BOOL  := 0;
  END_VAR
  IF NOT RESET AND tock = NOT TICK THEN
      Data[j]   := IN1;
      Data[j+1] := IN2;
      Data[j+2] := IN3;
      Data[j+3] := IN4;
      Data[j+4] := IN5;
      j := j + 5;
      tock := TICK;
  ELSE
      j := 1;
      tock := 0;
  END_IF;
  Finished := (j > 15);
END_FUNCTION_BLOCK

PROGRAM Boiler
  VAR
    Data  : ARRAY[1..15] OF BOOL;
    Ready : BOOL;
    CollectInput : F_CollectInput;
  END_VAR
  VAR
    TICK     AT %IX1.0 : BOOL;
    IN1      AT %IX0.3 : BOOL;
    IN2      AT %IX0.4 : BOOL;
    IN3      AT %IX0.5 : BOOL;
    IN4      AT %IX0.6 : BOOL;
    IN5      AT %IX0.7 : BOOL;
    OutReady AT %QX0.0 : BOOL := FALSE;
    FeedNext AT %QX0.1 : BOOL := FALSE;
    Out      AT %QX0.2 : BOOL;
  END_VAR
  CollectInput(TICK:=TICK, IN1:=IN1, IN2:=IN2, IN3:=IN3, IN4:=IN4, IN5:=IN5);
  Ready := CollectInput.Finished;
  FeedNext := 1;
  IF Ready THEN
    Out := (((((((((NOT (((NOT D[5]) AND (NOT D[2])) AND (NOT D[1]))) OR D[4]) AND ((NOT ((D[5] AND (NOT D[2])) AND (NOT D[1]))) OR D[3])) AND ((NOT (((NOT D[5]) AND D[2]) AND (NOT D[1]))) OR D[6])) AND ((NOT ((D[5] AND D[2]) AND (NOT D[1]))) OR D[7])) AND ((NOT (((NOT D[5]) AND (NOT D[2])) AND D[1])) OR D[8])) AND ((NOT ((D[5] AND (NOT D[2])) AND D[1])) OR D[10])) AND ((NOT (((NOT D[5]) AND D[2]) AND D[1])) OR D[9])) AND ((NOT ((D[5] AND D[2]) AND D[1])) OR D[11]));
    OutReady := 1;
    CollectInput(RESET:=TRUE);
  END_IF;
END_PROGRAM

CONFIGURATION Config0
  RESOURCE Res0 ON PLC
    TASK task0(INTERVAL := T#20ms,PRIORITY := 0);
    PROGRAM instance0 WITH task0 : Boiler;
  END_RESOURCE
END_CONFIGURATION

(* ---- 3-MUX_augur-aleph-tiers.st ---- *)
(*
This code implements a shuffled multiplexer with 3 control bits.
The control bits are: Data[1], Data[2], Data[10]
The input bits are: Data[4], Data[5], Data[3], Data[8], Data[6], Data[7], Data[11], Data[9]

The symbolic expression is:
(((((((~((~(D[1]) & ~(D[2])) & ~(D[10])) | D[4]) & (~((D[1] & ~(D[2])) & ~(D[10])) | D[5])) & (~((~(D[1]) & D[2]) & ~(D[10])) | D[3])) & (~((D[1] & D[2]) & ~(D[10])) | D[8])) & (~((~(D[1]) & ~(D[2])) & D[10]) | D[6])) & (~((D[1] & ~(D[2])) & D[10]) | D[7])) & (~((~(D[1]) & D[2]) & D[10]) | D[11])) & (~((D[1] & D[2]) & D[10]) | D[9])

*)

FUNCTION_BLOCK F_CollectInput
  VAR_IN_OUT
      Data : ARRAY[1..15] OF BOOL;
  END_VAR
  VAR_INPUT
      TICK  : BOOL := 0;
      IN1   : BOOL := 0;
      IN2   : BOOL := 0;
      IN3   : BOOL := 0;
      IN4   : BOOL := 0;
      IN5   : BOOL := 0;
      RESET : BOOL := FALSE;
  END_VAR
  VAR_OUTPUT
      Finished : BOOL;
  END_VAR
  VAR
      j    : USINT := 1;
      tock : BOOL  := 0;
  END_VAR
  IF NOT RESET AND tock = NOT TICK THEN
      Data[j]   := IN1;
      Data[j+1] := IN2;
      Data[j+2] := IN3;
      Data[j+3] := IN4;
      Data[j+4] := IN5;
      j := j + 5;
      tock := TICK;
  ELSE
      j := 1;
      tock := 0;
  END_IF;
  Finished := (j > 15);
END_FUNCTION_BLOCK

PROGRAM Boiler
  VAR
    Data  : ARRAY[1..15] OF BOOL;
    Ready : BOOL;
    CollectInput : F_CollectInput;
  END_VAR
  VAR
    TICK     AT %IX1.0 : BOOL;
    IN1      AT %IX0.3 : BOOL;
    IN2      AT %IX0.4 : BOOL;
    IN3      AT %IX0.5 : BOOL;
    IN4      AT %IX0.6 : BOOL;
    IN5      AT %IX0.7 : BOOL;
    OutReady AT %QX0.0 : BOOL := FALSE;
    FeedNext AT %QX0.1 : BOOL := FALSE;
    Out      AT %QX0.2 : BOOL;
  END_VAR
  CollectInput(TICK:=TICK, IN1:=IN1, IN2:=IN2, IN3:=IN3, IN4:=IN4, IN5:=IN5);
  Ready := CollectInput.Finished;
  FeedNext := 1;
  IF Ready THEN
    Out := (((((((((NOT (((NOT D[1]) AND (NOT D[2])) AND (NOT D[10]))) OR D[4]) AND ((NOT ((D[1] AND (NOT D[2])) AND (NOT D[10]))) OR D[5])) AND ((NOT (((NOT D[1]) AND D[2]) AND (NOT D[10]))) OR D[3])) AND ((NOT ((D[1] AND D[2]) AND (NOT D[10]))) OR D[8])) AND ((NOT (((NOT D[1]) AND (NOT D[2])) AND D[10])) OR D[6])) AND ((NOT ((D[1] AND (NOT D[2])) AND D[10])) OR D[7])) AND ((NOT (((NOT D[1]) AND D[2]) AND D[10])) OR D[11])) AND ((NOT ((D[1] AND D[2]) AND D[10])) OR D[9]));
    OutReady := 1;
    CollectInput(RESET:=TRUE);
  END_IF;
END_PROGRAM

CONFIGURATION Config0
  RESOURCE Res0 ON PLC
    TASK task0(INTERVAL := T#20ms,PRIORITY := 0);
    PROGRAM instance0 WITH task0 : Boiler;
  END_RESOURCE
END_CONFIGURATION

(* ---- 3-MUX_avert-munge-biggy.st ---- *)
(*
This code implements a shuffled multiplexer with 3 control bits.
The control bits are: Data[1], Data[2], Data[4]
The input bits are: Data[5], Data[3], Data[7], Data[6], Data[8], Data[9], Data[11], Data[10]

The symbolic expression is:
(((((((~((~(D[1]) & ~(D[2])) & ~(D[4])) | D[5]) & (~((D[1] & ~(D[2])) & ~(D[4])) | D[3])) & (~((~(D[1]) & D[2]) & ~(D[4])) | D[7])) & (~((D[1] & D[2]) & ~(D[4])) | D[6])) & (~((~(D[1]) & ~(D[2])) & D[4]) | D[8])) & (~((D[1] & ~(D[2])) & D[4]) | D[9])) & (~((~(D[1]) & D[2]) & D[4]) | D[11])) & (~((D[1] & D[2]) & D[4]) | D[10])

*)

FUNCTION_BLOCK F_CollectInput
  VAR_IN_OUT
      Data : ARRAY[1..15] OF BOOL;
  END_VAR
  VAR_INPUT
      TICK  : BOOL := 0;
      IN1   : BOOL := 0;
      IN2   : BOOL := 0;
      IN3   : BOOL := 0;
      IN4   : BOOL := 0;
      IN5   : BOOL := 0;
      RESET : BOOL := FALSE;
  END_VAR
  VAR_OUTPUT
      Finished : BOOL;
  END_VAR
  VAR
      j    : USINT := 1;
      tock : BOOL  := 0;
  END_VAR
  IF NOT RESET AND tock = NOT TICK THEN
      Data[j]   := IN1;
      Data[j+1] := IN2;
      Data[j+2] := IN3;
      Data[j+3] := IN4;
      Data[j+4] := IN5;
      j := j + 5;
      tock := TICK;
  ELSE
      j := 1;
      tock := 0;
  END_IF;
  Finished := (j > 15);
END_FUNCTION_BLOCK

PROGRAM Boiler
  VAR
    Data  : ARRAY[1..15] OF BOOL;
    Ready : BOOL;
    CollectInput : F_CollectInput;
  END_VAR
  VAR
    TICK     AT %IX1.0 : BOOL;
    IN1      AT %IX0.3 : BOOL;
    IN2      AT %IX0.4 : BOOL;
    IN3      AT %IX0.5 : BOOL;
    IN4      AT %IX0.6 : BOOL;
    IN5      AT %IX0.7 : BOOL;
    OutReady AT %QX0.0 : BOOL := FALSE;
    FeedNext AT %QX0.1 : BOOL := FALSE;
    Out      AT %QX0.2 : BOOL;
  END_VAR
  CollectInput(TICK:=TICK, IN1:=IN1, IN2:=IN2, IN3:=IN3, IN4:=IN4, IN5:=IN5);
  Ready := CollectInput.Finished;
  FeedNext := 1;
  IF Ready THEN
    Out := (((((((((NOT (((NOT D[1]) AND (NOT D[2])) AND (NOT D[4]))) OR D[5]) AND ((NOT ((D[1] AND (NOT D[2])) AND (NOT D[4]))) OR D[3])) AND ((NOT (((NOT D[1]) AND D[2]) AND (NOT D[4]))) OR D[7])) AND ((NOT ((D[1] AND D[2]) AND (NOT D[4]))) OR D[6])) AND ((NOT (((NOT D[1]) AND (NOT D[2])) AND D[4])) OR D[8])) AND ((NOT ((D[1] AND (NOT D[2])) AND D[4])) OR D[9])) AND ((NOT (((NOT D[1]) AND D[2]) AND D[4])) OR D[11])) AND ((NOT ((D[1] AND D[2]) AND D[4])) OR D[10]));
    OutReady := 1;
    CollectInput(RESET:=TRUE);
  END_IF;
END_PROGRAM

CONFIGURATION Config0
  RESOURCE Res0 ON PLC
    TASK task0(INTERVAL := T#20ms,PRIORITY := 0);
    PROGRAM instance0 WITH task0 : Boiler;
  END_RESOURCE
END_CONFIGURATION

(* ---- 3-MUX_being-wiper-plena.st ---- *)
(*
This code implements a shuffled multiplexer with 3 control bits.
The control bits are: Data[4], Data[2], Data[1]
The input bits are: Data[3], Data[8], Data[6], Data[7], Data[10], Data[11], Data[5], Data[9]

The symbolic expression is:
(((((((~((~(D[4]) & ~(D[2])) & ~(D[1])) | D[3]) & (~((D[4] & ~(D[2])) & ~(D[1])) | D[8])) & (~((~(D[4]) & D[2]) & ~(D[1])) | D[6])) & (~((D[4] & D[2]) & ~(D[1])) | D[7])) & (~((~(D[4]) & ~(D[2])) & D[1]) | D[10])) & (~((D[4] & ~(D[2])) & D[1]) | D[11])) & (~((~(D[4]) & D[2]) & D[1]) | D[5])) & (~((D[4] & D[2]) & D[1]) | D[9])

*)

FUNCTION_BLOCK F_CollectInput
  VAR_IN_OUT
      Data : ARRAY[1..15] OF BOOL;
  END_VAR
  VAR_INPUT
      TICK  : BOOL := 0;
      IN1   : BOOL := 0;
      IN2   : BOOL := 0;
      IN3   : BOOL := 0;
      IN4   : BOOL := 0;
      IN5   : BOOL := 0;
      RESET : BOOL := FALSE;
  END_VAR
  VAR_OUTPUT
      Finished : BOOL;
  END_VAR
  VAR
      j    : USINT := 1;
      tock : BOOL  := 0;
  END_VAR
  IF NOT RESET AND tock = NOT TICK THEN
      Data[j]   := IN1;
      Data[j+1] := IN2;
      Data[j+2] := IN3;
      Data[j+3] := IN4;
      Data[j+4] := IN5;
      j := j + 5;
      tock := TICK;
  ELSE
      j := 1;
      tock := 0;
  END_IF;
  Finished := (j > 15);
END_FUNCTION_BLOCK

PROGRAM Boiler
  VAR
    Data  : ARRAY[1..15] OF BOOL;
    Ready : BOOL;
    CollectInput : F_CollectInput;
  END_VAR
  VAR
    TICK     AT %IX1.0 : BOOL;
    IN1      AT %IX0.3 : BOOL;
    IN2      AT %IX0.4 : BOOL;
    IN3      AT %IX0.5 : BOOL;
    IN4      AT %IX0.6 : BOOL;
    IN5      AT %IX0.7 : BOOL;
    OutReady AT %QX0.0 : BOOL := FALSE;
    FeedNext AT %QX0.1 : BOOL := FALSE;
    Out      AT %QX0.2 : BOOL;
  END_VAR
  CollectInput(TICK:=TICK, IN1:=IN1, IN2:=IN2, IN3:=IN3, IN4:=IN4, IN5:=IN5);
  Ready := CollectInput.Finished;
  FeedNext := 1;
  IF Ready THEN
    Out := (((((((((NOT (((NOT D[4]) AND (NOT D[2])) AND (NOT D[1]))) OR D[3]) AND ((NOT ((D[4] AND (NOT D[2])) AND (NOT D[1]))) OR D[8])) AND ((NOT (((NOT D[4]) AND D[2]) AND (NOT D[1]))) OR D[6])) AND ((NOT ((D[4] AND D[2]) AND (NOT D[1]))) OR D[7])) AND ((NOT (((NOT D[4]) AND (NOT D[2])) AND D[1])) OR D[10])) AND ((NOT ((D[4] AND (NOT D[2])) AND D[1])) OR D[11])) AND ((NOT (((NOT D[4]) AND D[2]) AND D[1])) OR D[5])) AND ((NOT ((D[4] AND D[2]) AND D[1])) OR D[9]));
    OutReady := 1;
    CollectInput(RESET:=TRUE);
  END_IF;
END_PROGRAM

CONFIGURATION Config0
  RESOURCE Res0 ON PLC
    TASK task0(INTERVAL := T#20ms,PRIORITY := 0);
    PROGRAM instance0 WITH task0 : Boiler;
  END_RESOURCE
END_CONFIGURATION

(* ---- 3-MUX_blimp-folks-kilty.st ---- *)
(*
This code implements a shuffled multiplexer with 3 control bits.
The control bits are: Data[7], Data[2], Data[10]
The input bits are: Data[3], Data[1], Data[4], Data[6], Data[5], Data[8], Data[9], Data[11]

The symbolic expression is:
(((((((~((~(D[7]) & ~(D[2])) & ~(D[10])) | D[3]) & (~((D[7] & ~(D[2])) & ~(D[10])) | D[1])) & (~((~(D[7]) & D[2]) & ~(D[10])) | D[4])) & (~((D[7] & D[2]) & ~(D[10])) | D[6])) & (~((~(D[7]) & ~(D[2])) & D[10]) | D[5])) & (~((D[7] & ~(D[2])) & D[10]) | D[8])) & (~((~(D[7]) & D[2]) & D[10]) | D[9])) & (~((D[7] & D[2]) & D[10]) | D[11])

*)

FUNCTION_BLOCK F_CollectInput
  VAR_IN_OUT
      Data : ARRAY[1..15] OF BOOL;
  END_VAR
  VAR_INPUT
      TICK  : BOOL := 0;
      IN1   : BOOL := 0;
      IN2   : BOOL := 0;
      IN3   : BOOL := 0;
      IN4   : BOOL := 0;
      IN5   : BOOL := 0;
      RESET : BOOL := FALSE;
  END_VAR
  VAR_OUTPUT
      Finished : BOOL;
  END_VAR
  VAR
      j    : USINT := 1;
      tock : BOOL  := 0;
  END_VAR
  IF NOT RESET AND tock = NOT TICK THEN
      Data[j]   := IN1;
      Data[j+1] := IN2;
      Data[j+2] := IN3;
      Data[j+3] := IN4;
      Data[j+4] := IN5;
      j := j + 5;
      tock := TICK;
  ELSE
      j := 1;
      tock := 0;
  END_IF;
  Finished := (j > 15);
END_FUNCTION_BLOCK

PROGRAM Boiler
  VAR
    Data  : ARRAY[1..15] OF BOOL;
    Ready : BOOL;
    CollectInput : F_CollectInput;
  END_VAR
  VAR
    TICK     AT %IX1.0 : BOOL;
    IN1      AT %IX0.3 : BOOL;
    IN2      AT %IX0.4 : BOOL;
    IN3      AT %IX0.5 : BOOL;
    IN4      AT %IX0.6 : BOOL;
    IN5      AT %IX0.7 : BOOL;
    OutReady AT %QX0.0 : BOOL := FALSE;
    FeedNext AT %QX0.1 : BOOL := FALSE;
    Out      AT %QX0.2 : BOOL;
  END_VAR
  CollectInput(TICK:=TICK, IN1:=IN1, IN2:=IN2, IN3:=IN3, IN4:=IN4, IN5:=IN5);
  Ready := CollectInput.Finished;
  FeedNext := 1;
  IF Ready THEN
    Out := (((((((((NOT (((NOT D[7]) AND (NOT D[2])) AND (NOT D[10]))) OR D[3]) AND ((NOT ((D[7] AND (NOT D[2])) AND (NOT D[10]))) OR D[1])) AND ((NOT (((NOT D[7]) AND D[2]) AND (NOT D[10]))) OR D[4])) AND ((NOT ((D[7] AND D[2]) AND (NOT D[10]))) OR D[6])) AND ((NOT (((NOT D[7]) AND (NOT D[2])) AND D[10])) OR D[5])) AND ((NOT ((D[7] AND (NOT D[2])) AND D[10])) OR D[8])) AND ((NOT (((NOT D[7]) AND D[2]) AND D[10])) OR D[9])) AND ((NOT ((D[7] AND D[2]) AND D[10])) OR D[11]));
    OutReady := 1;
    CollectInput(RESET:=TRUE);
  END_IF;
END_PROGRAM

CONFIGURATION Config0
  RESOURCE Res0 ON PLC
    TASK task0(INTERVAL := T#20ms,PRIORITY := 0);
    PROGRAM instance0 WITH task0 : Boiler;
  END_RESOURCE
END_CONFIGURATION

(* ---- 3-MUX_brick-jings-relay.st ---- *)
(*
This code implements a shuffled multiplexer with 3 control bits.
The control bits are: Data[1], Data[3], Data[2]
The input bits are: Data[4], Data[6], Data[7], Data[5], Data[8], Data[10], Data[11], Data[9]

The symbolic expression is:
(((((((~((~(D[1]) & ~(D[3])) & ~(D[2])) | D[4]) & (~((D[1] & ~(D[3])) & ~(D[2])) | D[6])) & (~((~(D[1]) & D[3]) & ~(D[2])) | D[7])) & (~((D[1] & D[3]) & ~(D[2])) | D[5])) & (~((~(D[1]) & ~(D[3])) & D[2]) | D[8])) & (~((D[1] & ~(D[3])) & D[2]) | D[10])) & (~((~(D[1]) & D[3]) & D[2]) | D[11])) & (~((D[1] & D[3]) & D[2]) | D[9])

*)

FUNCTION_BLOCK F_CollectInput
  VAR_IN_OUT
      Data : ARRAY[1..15] OF BOOL;
  END_VAR
  VAR_INPUT
      TICK  : BOOL := 0;
      IN1   : BOOL := 0;
      IN2   : BOOL := 0;
      IN3   : BOOL := 0;
      IN4   : BOOL := 0;
      IN5   : BOOL := 0;
      RESET : BOOL := FALSE;
  END_VAR
  VAR_OUTPUT
      Finished : BOOL;
  END_VAR
  VAR
      j    : USINT := 1;
      tock : BOOL  := 0;
  END_VAR
  IF NOT RESET AND tock = NOT TICK THEN
      Data[j]   := IN1;
      Data[j+1] := IN2;
      Data[j+2] := IN3;
      Data[j+3] := IN4;
      Data[j+4] := IN5;
      j := j + 5;
      tock := TICK;
  ELSE
      j := 1;
      tock := 0;
  END_IF;
  Finished := (j > 15);
END_FUNCTION_BLOCK

PROGRAM Boiler
  VAR
    Data  : ARRAY[1..15] OF BOOL;
    Ready : BOOL;
    CollectInput : F_CollectInput;
  END_VAR
  VAR
    TICK     AT %IX1.0 : BOOL;
    IN1      AT %IX0.3 : BOOL;
    IN2      AT %IX0.4 : BOOL;
    IN3      AT %IX0.5 : BOOL;
    IN4      AT %IX0.6 : BOOL;
    IN5      AT %IX0.7 : BOOL;
    OutReady AT %QX0.0 : BOOL := FALSE;
    FeedNext AT %QX0.1 : BOOL := FALSE;
    Out      AT %QX0.2 : BOOL;
  END_VAR
  CollectInput(TICK:=TICK, IN1:=IN1, IN2:=IN2, IN3:=IN3, IN4:=IN4, IN5:=IN5);
  Ready := CollectInput.Finished;
  FeedNext := 1;
  IF Ready THEN
    Out := (((((((((NOT (((NOT D[1]) AND (NOT D[3])) AND (NOT D[2]))) OR D[4]) AND ((NOT ((D[1] AND (NOT D[3])) AND (NOT D[2]))) OR D[6])) AND ((NOT (((NOT D[1]) AND D[3]) AND (NOT D[2]))) OR D[7])) AND ((NOT ((D[1] AND D[3]) AND (NOT D[2]))) OR D[5])) AND ((NOT (((NOT D[1]) AND (NOT D[3])) AND D[2])) OR D[8])) AND ((NOT ((D[1] AND (NOT D[3])) AND D[2])) OR D[10])) AND ((NOT (((NOT D[1]) AND D[3]) AND D[2])) OR D[11])) AND ((NOT ((D[1] AND D[3]) AND D[2])) OR D[9]));
    OutReady := 1;
    CollectInput(RESET:=TRUE);
  END_IF;
END_PROGRAM

CONFIGURATION Config0
  RESOURCE Res0 ON PLC
    TASK task0(INTERVAL := T#20ms,PRIORITY := 0);
    PROGRAM instance0 WITH task0 : Boiler;
  END_RESOURCE
END_CONFIGURATION

(* ---- 3-MUX_brood-tuxes-dotes.st ---- *)
(*
This code implements a shuffled multiplexer with 3 control bits.
The control bits are: Data[1], Data[2], Data[3]
The input bits are: Data[5], Data[4], Data[8], Data[10], Data[6], Data[9], Data[7], Data[11]

The symbolic expression is:
(((((((~((~(D[1]) & ~(D[2])) & ~(D[3])) | D[5]) & (~((D[1] & ~(D[2])) & ~(D[3])) | D[4])) & (~((~(D[1]) & D[2]) & ~(D[3])) | D[8])) & (~((D[1] & D[2]) & ~(D[3])) | D[10])) & (~((~(D[1]) & ~(D[2])) & D[3]) | D[6])) & (~((D[1] & ~(D[2])) & D[3]) | D[9])) & (~((~(D[1]) & D[2]) & D[3]) | D[7])) & (~((D[1] & D[2]) & D[3]) | D[11])

*)

FUNCTION_BLOCK F_CollectInput
  VAR_IN_OUT
      Data : ARRAY[1..15] OF BOOL;
  END_VAR
  VAR_INPUT
      TICK  : BOOL := 0;
      IN1   : BOOL := 0;
      IN2   : BOOL := 0;
      IN3   : BOOL := 0;
      IN4   : BOOL := 0;
      IN5   : BOOL := 0;
      RESET : BOOL := FALSE;
  END_VAR
  VAR_OUTPUT
      Finished : BOOL;
  END_VAR
  VAR
      j    : USINT := 1;
      tock : BOOL  := 0;
  END_VAR
  IF NOT RESET AND tock = NOT TICK THEN
      Data[j]   := IN1;
      Data[j+1] := IN2;
      Data[j+2] := IN3;
      Data[j+3] := IN4;
      Data[j+4] := IN5;
      j := j + 5;
      tock := TICK;
  ELSE
      j := 1;
      tock := 0;
  END_IF;
  Finished := (j > 15);
END_FUNCTION_BLOCK

PROGRAM Boiler
  VAR
    Data  : ARRAY[1..15] OF BOOL;
    Ready : BOOL;
    CollectInput : F_CollectInput;
  END_VAR
  VAR
    TICK     AT %IX1.0 : BOOL;
    IN1      AT %IX0.3 : BOOL;
    IN2      AT %IX0.4 : BOOL;
    IN3      AT %IX0.5 : BOOL;
    IN4      AT %IX0.6 : BOOL;
    IN5      AT %IX0.7 : BOOL;
    OutReady AT %QX0.0 : BOOL := FALSE;
    FeedNext AT %QX0.1 : BOOL := FALSE;
    Out      AT %QX0.2 : BOOL;
  END_VAR
  CollectInput(TICK:=TICK, IN1:=IN1, IN2:=IN2, IN3:=IN3, IN4:=IN4, IN5:=IN5);
  Ready := CollectInput.Finished;
  FeedNext := 1;
  IF Ready THEN
    Out := (((((((((NOT (((NOT D[1]) AND (NOT D[2])) AND (NOT D[3]))) OR D[5]) AND ((NOT ((D[1] AND (NOT D[2])) AND (NOT D[3]))) OR D[4])) AND ((NOT (((NOT D[1]) AND D[2]) AND (NOT D[3]))) OR D[8])) AND ((NOT ((D[1] AND D[2]) AND (NOT D[3]))) OR D[10])) AND ((NOT (((NOT D[1]) AND (NOT D[2])) AND D[3])) OR D[6])) AND ((NOT ((D[1] AND (NOT D[2])) AND D[3])) OR D[9])) AND ((NOT (((NOT D[1]) AND D[2]) AND D[3])) OR D[7])) AND ((NOT ((D[1] AND D[2]) AND D[3])) OR D[11]));
    OutReady := 1;
    CollectInput(RESET:=TRUE);
  END_IF;
END_PROGRAM

CONFIGURATION Config0
  RESOURCE Res0 ON PLC
    TASK task0(INTERVAL := T#20ms,PRIORITY := 0);
    PROGRAM instance0 WITH task0 : Boiler;
  END_RESOURCE
END_CONFIGURATION

(* ---- 3-MUX_bunco-towed-supra.st ---- *)
(*
This code implements a shuffled multiplexer with 3 control bits.
The control bits are: Data[4], Data[1], Data[3]
The input bits are: Data[2], Data[5], Data[6], Data[7], Data[8], Data[10], Data[9], Data[11]

The symbolic expression is:
(((((((~((~(D[4]) & ~(D[1])) & ~(D[3])) | D[2]) & (~((D[4] & ~(D[1])) & ~(D[3])) | D[5])) & (~((~(D[4]) & D[1]) & ~(D[3])) | D[6])) & (~((D[4] & D[1]) & ~(D[3])) | D[7])) & (~((~(D[4]) & ~(D[1])) & D[3]) | D[8])) & (~((D[4] & ~(D[1])) & D[3]) | D[10])) & (~((~(D[4]) & D[1]) & D[3]) | D[9])) & (~((D[4] & D[1]) & D[3]) | D[11])

*)

FUNCTION_BLOCK F_CollectInput
  VAR_IN_OUT
      Data : ARRAY[1..15] OF BOOL;
  END_VAR
  VAR_INPUT
      TICK  : BOOL := 0;
      IN1   : BOOL := 0;
      IN2   : BOOL := 0;
      IN3   : BOOL := 0;
      IN4   : BOOL := 0;
      IN5   : BOOL := 0;
      RESET : BOOL := FALSE;
  END_VAR
  VAR_OUTPUT
      Finished : BOOL;
  END_VAR
  VAR
      j    : USINT := 1;
      tock : BOOL  := 0;
  END_VAR
  IF NOT RESET AND tock = NOT TICK THEN
      Data[j]   := IN1;
      Data[j+1] := IN2;
      Data[j+2] := IN3;
      Data[j+3] := IN4;
      Data[j+4] := IN5;
      j := j + 5;
      tock := TICK;
  ELSE
      j := 1;
      tock := 0;
  END_IF;
  Finished := (j > 15);
END_FUNCTION_BLOCK

PROGRAM Boiler
  VAR
    Data  : ARRAY[1..15] OF BOOL;
    Ready : BOOL;
    CollectInput : F_CollectInput;
  END_VAR
  VAR
    TICK     AT %IX1.0 : BOOL;
    IN1      AT %IX0.3 : BOOL;
    IN2      AT %IX0.4 : BOOL;
    IN3      AT %IX0.5 : BOOL;
    IN4      AT %IX0.6 : BOOL;
    IN5      AT %IX0.7 : BOOL;
    OutReady AT %QX0.0 : BOOL := FALSE;
    FeedNext AT %QX0.1 : BOOL := FALSE;
    Out      AT %QX0.2 : BOOL;
  END_VAR
  CollectInput(TICK:=TICK, IN1:=IN1, IN2:=IN2, IN3:=IN3, IN4:=IN4, IN5:=IN5);
  Ready := CollectInput.Finished;
  FeedNext := 1;
  IF Ready THEN
    Out := (((((((((NOT (((NOT D[4]) AND (NOT D[1])) AND (NOT D[3]))) OR D[2]) AND ((NOT ((D[4] AND (NOT D[1])) AND (NOT D[3]))) OR D[5])) AND ((NOT (((NOT D[4]) AND D[1]) AND (NOT D[3]))) OR D[6])) AND ((NOT ((D[4] AND D[1]) AND (NOT D[3]))) OR D[7])) AND ((NOT (((NOT D[4]) AND (NOT D[1])) AND D[3])) OR D[8])) AND ((NOT ((D[4] AND (NOT D[1])) AND D[3])) OR D[10])) AND ((NOT (((NOT D[4]) AND D[1]) AND D[3])) OR D[9])) AND ((NOT ((D[4] AND D[1]) AND D[3])) OR D[11]));
    OutReady := 1;
    CollectInput(RESET:=TRUE);
  END_IF;
END_PROGRAM

CONFIGURATION Config0
  RESOURCE Res0 ON PLC
    TASK task0(INTERVAL := T#20ms,PRIORITY := 0);
    PROGRAM instance0 WITH task0 : Boiler;
  END_RESOURCE
END_CONFIGURATION

(* ---- 3-MUX_cauls-phony-gnats.st ---- *)
(*
This code implements a shuffled multiplexer with 3 control bits.
The control bits are: Data[6], Data[3], Data[1]
The input bits are: Data[4], Data[2], Data[7], Data[8], Data[9], Data[10], Data[11], Data[5]

The symbolic expression is:
(((((((~((~(D[6]) & ~(D[3])) & ~(D[1])) | D[4]) & (~((D[6] & ~(D[3])) & ~(D[1])) | D[2])) & (~((~(D[6]) & D[3]) & ~(D[1])) | D[7])) & (~((D[6] & D[3]) & ~(D[1])) | D[8])) & (~((~(D[6]) & ~(D[3])) & D[1]) | D[9])) & (~((D[6] & ~(D[3])) & D[1]) | D[10])) & (~((~(D[6]) & D[3]) & D[1]) | D[11])) & (~((D[6] & D[3]) & D[1]) | D[5])

*)

FUNCTION_BLOCK F_CollectInput
  VAR_IN_OUT
      Data : ARRAY[1..15] OF BOOL;
  END_VAR
  VAR_INPUT
      TICK  : BOOL := 0;
      IN1   : BOOL := 0;
      IN2   : BOOL := 0;
      IN3   : BOOL := 0;
      IN4   : BOOL := 0;
      IN5   : BOOL := 0;
      RESET : BOOL := FALSE;
  END_VAR
  VAR_OUTPUT
      Finished : BOOL;
  END_VAR
  VAR
      j    : USINT := 1;
      tock : BOOL  := 0;
  END_VAR
  IF NOT RESET AND tock = NOT TICK THEN
      Data[j]   := IN1;
      Data[j+1] := IN2;
      Data[j+2] := IN3;
      Data[j+3] := IN4;
      Data[j+4] := IN5;
      j := j + 5;
      tock := TICK;
  ELSE
      j := 1;
      tock := 0;
  END_IF;
  Finished := (j > 15);
END_FUNCTION_BLOCK

PROGRAM Boiler
  VAR
    Data  : ARRAY[1..15] OF BOOL;
    Ready : BOOL;
    CollectInput : F_CollectInput;
  END_VAR
  VAR
    TICK     AT %IX1.0 : BOOL;
    IN1      AT %IX0.3 : BOOL;
    IN2      AT %IX0.4 : BOOL;
    IN3      AT %IX0.5 : BOOL;
    IN4      AT %IX0.6 : BOOL;
    IN5      AT %IX0.7 : BOOL;
    OutReady AT %QX0.0 : BOOL := FALSE;
    FeedNext AT %QX0.1 : BOOL := FALSE;
    Out      AT %QX0.2 : BOOL;
  END_VAR
  CollectInput(TICK:=TICK, IN1:=IN1, IN2:=IN2, IN3:=IN3, IN4:=IN4, IN5:=IN5);
  Ready := CollectInput.Finished;
  FeedNext := 1;
  IF Ready THEN
    Out := (((((((((NOT (((NOT D[6]) AND (NOT D[3])) AND (NOT D[1]))) OR D[4]) AND ((NOT ((D[6] AND (NOT D[3])) AND (NOT D[1]))) OR D[2])) AND ((NOT (((NOT D[6]) AND D[3]) AND (NOT D[1]))) OR D[7])) AND ((NOT ((D[6] AND D[3]) AND (NOT D[1]))) OR D[8])) AND ((NOT (((NOT D[6]) AND (NOT D[3])) AND D[1])) OR D[9])) AND ((NOT ((D[6] AND (NOT D[3])) AND D[1])) OR D[10])) AND ((NOT (((NOT D[6]) AND D[3]) AND D[1])) OR D[11])) AND ((NOT ((D[6] AND D[3]) AND D[1])) OR D[5]));
    OutReady := 1;
    CollectInput(RESET:=TRUE);
  END_IF;
END_PROGRAM

CONFIGURATION Config0
  RESOURCE Res0 ON PLC
    TASK task0(INTERVAL := T#20ms,PRIORITY := 0);
    PROGRAM instance0 WITH task0 : Boiler;
  END_RESOURCE
END_CONFIGURATION

(* ---- 3-MUX_ceded-muser-treys.st ---- *)
(*
This code implements a shuffled multiplexer with 3 control bits.
The control bits are: Data[1], Data[5], Data[2]
The input bits are: Data[4], Data[3], Data[6], Data[7], Data[9], Data[8], Data[11], Data[10]

The symbolic expression is:
(((((((~((~(D[1]) & ~(D[5])) & ~(D[2])) | D[4]) & (~((D[1] & ~(D[5])) & ~(D[2])) | D[3])) & (~((~(D[1]) & D[5]) & ~(D[2])) | D[6])) & (~((D[1] & D[5]) & ~(D[2])) | D[7])) & (~((~(D[1]) & ~(D[5])) & D[2]) | D[9])) & (~((D[1] & ~(D[5])) & D[2]) | D[8])) & (~((~(D[1]) & D[5]) & D[2]) | D[11])) & (~((D[1] & D[5]) & D[2]) | D[10])

*)

FUNCTION_BLOCK F_CollectInput
  VAR_IN_OUT
      Data : ARRAY[1..15] OF BOOL;
  END_VAR
  VAR_INPUT
      TICK  : BOOL := 0;
      IN1   : BOOL := 0;
      IN2   : BOOL := 0;
      IN3   : BOOL := 0;
      IN4   : BOOL := 0;
      IN5   : BOOL := 0;
      RESET : BOOL := FALSE;
  END_VAR
  VAR_OUTPUT
      Finished : BOOL;
  END_VAR
  VAR
      j    : USINT := 1;
      tock : BOOL  := 0;
  END_VAR
  IF NOT RESET AND tock = NOT TICK THEN
      Data[j]   := IN1;
      Data[j+1] := IN2;
      Data[j+2] := IN3;
      Data[j+3] := IN4;
      Data[j+4] := IN5;
      j := j + 5;
      tock := TICK;
  ELSE
      j := 1;
      tock := 0;
  END_IF;
  Finished := (j > 15);
END_FUNCTION_BLOCK

PROGRAM Boiler
  VAR
    Data  : ARRAY[1..15] OF BOOL;
    Ready : BOOL;
    CollectInput : F_CollectInput;
  END_VAR
  VAR
    TICK     AT %IX1.0 : BOOL;
    IN1      AT %IX0.3 : BOOL;
    IN2      AT %IX0.4 : BOOL;
    IN3      AT %IX0.5 : BOOL;
    IN4      AT %IX0.6 : BOOL;
    IN5      AT %IX0.7 : BOOL;
    OutReady AT %QX0.0 : BOOL := FALSE;
    FeedNext AT %QX0.1 : BOOL := FALSE;
    Out      AT %QX0.2 : BOOL;
  END_VAR
  CollectInput(TICK:=TICK, IN1:=IN1, IN2:=IN2, IN3:=IN3, IN4:=IN4, IN5:=IN5);
  Ready := CollectInput.Finished;
  FeedNext := 1;
  IF Ready THEN
    Out := (((((((((NOT (((NOT D[1]) AND (NOT D[5])) AND (NOT D[2]))) OR D[4]) AND ((NOT ((D[1] AND (NOT D[5])) AND (NOT D[2]))) OR D[3])) AND ((NOT (((NOT D[1]) AND D[5]) AND (NOT D[2]))) OR D[6])) AND ((NOT ((D[1] AND D[5]) AND (NOT D[2]))) OR D[7])) AND ((NOT (((NOT D[1]) AND (NOT D[5])) AND D[2])) OR D[9])) AND ((NOT ((D[1] AND (NOT D[5])) AND D[2])) OR D[8])) AND ((NOT (((NOT D[1]) AND D[5]) AND D[2])) OR D[11])) AND ((NOT ((D[1] AND D[5]) AND D[2])) OR D[10]));
    OutReady := 1;
    CollectInput(RESET:=TRUE);
  END_IF;
END_PROGRAM

CONFIGURATION Config0
  RESOURCE Res0 ON PLC
    TASK task0(INTERVAL := T#20ms,PRIORITY := 0);
    PROGRAM instance0 WITH task0 : Boiler;
  END_RESOURCE
END_CONFIGURATION

(* ---- 3-MUX_clues-cukes-smurf.st ---- *)
(*
This code implements a shuffled multiplexer with 3 control bits.
The control bits are: Data[2], Data[6], Data[4]
The input bits are: Data[1], Data[8], Data[3], Data[7], Data[5], Data[9], Data[10], Data[11]

The symbolic expression is:
(((((((~((~(D[2]) & ~(D[6])) & ~(D[4])) | D[1]) & (~((D[2] & ~(D[6])) & ~(D[4])) | D[8])) & (~((~(D[2]) & D[6]) & ~(D[4])) | D[3])) & (~((D[2] & D[6]) & ~(D[4])) | D[7])) & (~((~(D[2]) & ~(D[6])) & D[4]) | D[5])) & (~((D[2] & ~(D[6])) & D[4]) | D[9])) & (~((~(D[2]) & D[6]) & D[4]) | D[10])) & (~((D[2] & D[6]) & D[4]) | D[11])

*)

FUNCTION_BLOCK F_CollectInput
  VAR_IN_OUT
      Data : ARRAY[1..15] OF BOOL;
  END_VAR
  VAR_INPUT
      TICK  : BOOL := 0;
      IN1   : BOOL := 0;
      IN2   : BOOL := 0;
      IN3   : BOOL := 0;
      IN4   : BOOL := 0;
      IN5   : BOOL := 0;
      RESET : BOOL := FALSE;
  END_VAR
  VAR_OUTPUT
      Finished : BOOL;
  END_VAR
  VAR
      j    : USINT := 1;
      tock : BOOL  := 0;
  END_VAR
  IF NOT RESET AND tock = NOT TICK THEN
      Data[j]   := IN1;
      Data[j+1] := IN2;
      Data[j+2] := IN3;
      Data[j+3] := IN4;
      Data[j+4] := IN5;
      j := j + 5;
      tock := TICK;
  ELSE
      j := 1;
      tock := 0;
  END_IF;
  Finished := (j > 15);
END_FUNCTION_BLOCK

PROGRAM Boiler
  VAR
    Data  : ARRAY[1..15] OF BOOL;
    Ready : BOOL;
    CollectInput : F_CollectInput;
  END_VAR
  VAR
    TICK     AT %IX1.0 : BOOL;
    IN1      AT %IX0.3 : BOOL;
    IN2      AT %IX0.4 : BOOL;
    IN3      AT %IX0.5 : BOOL;
    IN4      AT %IX0.6 : BOOL;
    IN5      AT %IX0.7 : BOOL;
    OutReady AT %QX0.0 : BOOL := FALSE;
    FeedNext AT %QX0.1 : BOOL := FALSE;
    Out      AT %QX0.2 : BOOL;
  END_VAR
  CollectInput(TICK:=TICK, IN1:=IN1, IN2:=IN2, IN3:=IN3, IN4:=IN4, IN5:=IN5);
  Ready := CollectInput.Finished;
  FeedNext := 1;
  IF Ready THEN
    Out := (((((((((NOT (((NOT D[2]) AND (NOT D[6])) AND (NOT D[4]))) OR D[1]) AND ((NOT ((D[2] AND (NOT D[6])) AND (NOT D[4]))) OR D[8])) AND ((NOT (((NOT D[2]) AND D[6]) AND (NOT D[4]))) OR D[3])) AND ((NOT ((D[2] AND D[6]) AND (NOT D[4]))) OR D[7])) AND ((NOT (((NOT D[2]) AND (NOT D[6])) AND D[4])) OR D[5])) AND ((NOT ((D[2] AND (NOT D[6])) AND D[4])) OR D[9])) AND ((NOT (((NOT D[2]) AND D[6]) AND D[4])) OR D[10])) AND ((NOT ((D[2] AND D[6]) AND D[4])) OR D[11]));
    OutReady := 1;
    CollectInput(RESET:=TRUE);
  END_IF;
END_PROGRAM

CONFIGURATION Config0
  RESOURCE Res0 ON PLC
    TASK task0(INTERVAL := T#20ms,PRIORITY := 0);
    PROGRAM instance0 WITH task0 : Boiler;
  END_RESOURCE
END_CONFIGURATION

(* ---- 3-MUX_coals-oweth-gazer.st ---- *)
(*
This code implements a shuffled multiplexer with 3 control bits.
The control bits are: Data[2], Data[6], Data[1]
The input bits are: Data[3], Data[7], Data[4], Data[5], Data[8], Data[10], Data[9], Data[11]

The symbolic expression is:
(((((((~((~(D[2]) & ~(D[6])) & ~(D[1])) | D[3]) & (~((D[2] & ~(D[6])) & ~(D[1])) | D[7])) & (~((~(D[2]) & D[6]) & ~(D[1])) | D[4])) & (~((D[2] & D[6]) & ~(D[1])) | D[5])) & (~((~(D[2]) & ~(D[6])) & D[1]) | D[8])) & (~((D[2] & ~(D[6])) & D[1]) | D[10])) & (~((~(D[2]) & D[6]) & D[1]) | D[9])) & (~((D[2] & D[6]) & D[1]) | D[11])

*)

FUNCTION_BLOCK F_CollectInput
  VAR_IN_OUT
      Data : ARRAY[1..15] OF BOOL;
  END_VAR
  VAR_INPUT
      TICK  : BOOL := 0;
      IN1   : BOOL := 0;
      IN2   : BOOL := 0;
      IN3   : BOOL := 0;
      IN4   : BOOL := 0;
      IN5   : BOOL := 0;
      RESET : BOOL := FALSE;
  END_VAR
  VAR_OUTPUT
      Finished : BOOL;
  END_VAR
  VAR
      j    : USINT := 1;
      tock : BOOL  := 0;
  END_VAR
  IF NOT RESET AND tock = NOT TICK THEN
      Data[j]   := IN1;
      Data[j+1] := IN2;
      Data[j+2] := IN3;
      Data[j+3] := IN4;
      Data[j+4] := IN5;
      j := j + 5;
      tock := TICK;
  ELSE
      j := 1;
      tock := 0;
  END_IF;
  Finished := (j > 15);
END_FUNCTION_BLOCK

PROGRAM Boiler
  VAR
    Data  : ARRAY[1..15] OF BOOL;
    Ready : BOOL;
    CollectInput : F_CollectInput;
  END_VAR
  VAR
    TICK     AT %IX1.0 : BOOL;
    IN1      AT %IX0.3 : BOOL;
    IN2      AT %IX0.4 : BOOL;
    IN3      AT %IX0.5 : BOOL;
    IN4      AT %IX0.6 : BOOL;
    IN5      AT %IX0.7 : BOOL;
    OutReady AT %QX0.0 : BOOL := FALSE;
    FeedNext AT %QX0.1 : BOOL := FALSE;
    Out      AT %QX0.2 : BOOL;
  END_VAR
  CollectInput(TICK:=TICK, IN1:=IN1, IN2:=IN2, IN3:=IN3, IN4:=IN4, IN5:=IN5);
  Ready := CollectInput.Finished;
  FeedNext := 1;
  IF Ready THEN
    Out := (((((((((NOT (((NOT D[2]) AND (NOT D[6])) AND (NOT D[1]))) OR D[3]) AND ((NOT ((D[2] AND (NOT D[6])) AND (NOT D[1]))) OR D[7])) AND ((NOT (((NOT D[2]) AND D[6]) AND (NOT D[1]))) OR D[4])) AND ((NOT ((D[2] AND D[6]) AND (NOT D[1]))) OR D[5])) AND ((NOT (((NOT D[2]) AND (NOT D[6])) AND D[1])) OR D[8])) AND ((NOT ((D[2] AND (NOT D[6])) AND D[1])) OR D[10])) AND ((NOT (((NOT D[2]) AND D[6]) AND D[1])) OR D[9])) AND ((NOT ((D[2] AND D[6]) AND D[1])) OR D[11]));
    OutReady := 1;
    CollectInput(RESET:=TRUE);
  END_IF;
END_PROGRAM

CONFIGURATION Config0
  RESOURCE Res0 ON PLC
    TASK task0(INTERVAL := T#20ms,PRIORITY := 0);
    PROGRAM instance0 WITH task0 : Boiler;
  END_RESOURCE
END_CONFIGURATION

(* ---- 3-MUX_cress-paned-squib.st ---- *)
(*
This code implements a shuffled multiplexer with 3 control bits.
The control bits are: Data[5], Data[3], Data[1]
The input bits are: Data[2], Data[6], Data[4], Data[7], Data[8], Data[9], Data[10], Data[11]

The symbolic expression is:
(((((((~((~(D[5]) & ~(D[3])) & ~(D[1])) | D[2]) & (~((D[5] & ~(D[3])) & ~(D[1])) | D[6])) & (~((~(D[5]) & D[3]) & ~(D[1])) | D[4])) & (~((D[5] & D[3]) & ~(D[1])) | D[7])) & (~((~(D[5]) & ~(D[3])) & D[1]) | D[8])) & (~((D[5] & ~(D[3])) & D[1]) | D[9])) & (~((~(D[5]) & D[3]) & D[1]) | D[10])) & (~((D[5] & D[3]) & D[1]) | D[11])

*)

FUNCTION_BLOCK F_CollectInput
  VAR_IN_OUT
      Data : ARRAY[1..15] OF BOOL;
  END_VAR
  VAR_INPUT
      TICK  : BOOL := 0;
      IN1   : BOOL := 0;
      IN2   : BOOL := 0;
      IN3   : BOOL := 0;
      IN4   : BOOL := 0;
      IN5   : BOOL := 0;
      RESET : BOOL := FALSE;
  END_VAR
  VAR_OUTPUT
      Finished : BOOL;
  END_VAR
  VAR
      j    : USINT := 1;
      tock : BOOL  := 0;
  END_VAR
  IF NOT RESET AND tock = NOT TICK THEN
      Data[j]   := IN1;
      Data[j+1] := IN2;
      Data[j+2] := IN3;
      Data[j+3] := IN4;
      Data[j+4] := IN5;
      j := j + 5;
      tock := TICK;
  ELSE
      j := 1;
      tock := 0;
  END_IF;
  Finished := (j > 15);
END_FUNCTION_BLOCK

PROGRAM Boiler
  VAR
    Data  : ARRAY[1..15] OF BOOL;
    Ready : BOOL;
    CollectInput : F_CollectInput;
  END_VAR
  VAR
    TICK     AT %IX1.0 : BOOL;
    IN1      AT %IX0.3 : BOOL;
    IN2      AT %IX0.4 : BOOL;
    IN3      AT %IX0.5 : BOOL;
    IN4      AT %IX0.6 : BOOL;
    IN5      AT %IX0.7 : BOOL;
    OutReady AT %QX0.0 : BOOL := FALSE;
    FeedNext AT %QX0.1 : BOOL := FALSE;
    Out      AT %QX0.2 : BOOL;
  END_VAR
  CollectInput(TICK:=TICK, IN1:=IN1, IN2:=IN2, IN3:=IN3, IN4:=IN4, IN5:=IN5);
  Ready := CollectInput.Finished;
  FeedNext := 1;
  IF Ready THEN
    Out := (((((((((NOT (((NOT D[5]) AND (NOT D[3])) AND (NOT D[1]))) OR D[2]) AND ((NOT ((D[5] AND (NOT D[3])) AND (NOT D[1]))) OR D[6])) AND ((NOT (((NOT D[5]) AND D[3]) AND (NOT D[1]))) OR D[4])) AND ((NOT ((D[5] AND D[3]) AND (NOT D[1]))) OR D[7])) AND ((NOT (((NOT D[5]) AND (NOT D[3])) AND D[1])) OR D[8])) AND ((NOT ((D[5] AND (NOT D[3])) AND D[1])) OR D[9])) AND ((NOT (((NOT D[5]) AND D[3]) AND D[1])) OR D[10])) AND ((NOT ((D[5] AND D[3]) AND D[1])) OR D[11]));
    OutReady := 1;
    CollectInput(RESET:=TRUE);
  END_IF;
END_PROGRAM

CONFIGURATION Config0
  RESOURCE Res0 ON PLC
    TASK task0(INTERVAL := T#20ms,PRIORITY := 0);
    PROGRAM instance0 WITH task0 : Boiler;
  END_RESOURCE
END_CONFIGURATION

(* ---- 3-MUX_crude-fiver-copse.st ---- *)
(*
This code implements a shuffled multiplexer with 3 control bits.
The control bits are: Data[4], Data[3], Data[1]
The input bits are: Data[2], Data[6], Data[7], Data[5], Data[10], Data[8], Data[9], Data[11]

The symbolic expression is:
(((((((~((~(D[4]) & ~(D[3])) & ~(D[1])) | D[2]) & (~((D[4] & ~(D[3])) & ~(D[1])) | D[6])) & (~((~(D[4]) & D[3]) & ~(D[1])) | D[7])) & (~((D[4] & D[3]) & ~(D[1])) | D[5])) & (~((~(D[4]) & ~(D[3])) & D[1]) | D[10])) & (~((D[4] & ~(D[3])) & D[1]) | D[8])) & (~((~(D[4]) & D[3]) & D[1]) | D[9])) & (~((D[4] & D[3]) & D[1]) | D[11])

*)

FUNCTION_BLOCK F_CollectInput
  VAR_IN_OUT
      Data : ARRAY[1..15] OF BOOL;
  END_VAR
  VAR_INPUT
      TICK  : BOOL := 0;
      IN1   : BOOL := 0;
      IN2   : BOOL := 0;
      IN3   : BOOL := 0;
      IN4   : BOOL := 0;
      IN5   : BOOL := 0;
      RESET : BOOL := FALSE;
  END_VAR
  VAR_OUTPUT
      Finished : BOOL;
  END_VAR
  VAR
      j    : USINT := 1;
      tock : BOOL  := 0;
  END_VAR
  IF NOT RESET AND tock = NOT TICK THEN
      Data[j]   := IN1;
      Data[j+1] := IN2;
      Data[j+2] := IN3;
      Data[j+3] := IN4;
      Data[j+4] := IN5;
      j := j + 5;
      tock := TICK;
  ELSE
      j := 1;
      tock := 0;
  END_IF;
  Finished := (j > 15);
END_FUNCTION_BLOCK

PROGRAM Boiler
  VAR
    Data  : ARRAY[1..15] OF BOOL;
    Ready : BOOL;
    CollectInput : F_CollectInput;
  END_VAR
  VAR
    TICK     AT %IX1.0 : BOOL;
    IN1      AT %IX0.3 : BOOL;
    IN2      AT %IX0.4 : BOOL;
    IN3      AT %IX0.5 : BOOL;
    IN4      AT %IX0.6 : BOOL;
    IN5      AT %IX0.7 : BOOL;
    OutReady AT %QX0.0 : BOOL := FALSE;
    FeedNext AT %QX0.1 : BOOL := FALSE;
    Out      AT %QX0.2 : BOOL;
  END_VAR
  CollectInput(TICK:=TICK, IN1:=IN1, IN2:=IN2, IN3:=IN3, IN4:=IN4, IN5:=IN5);
  Ready := CollectInput.Finished;
  FeedNext := 1;
  IF Ready THEN
    Out := (((((((((NOT (((NOT D[4]) AND (NOT D[3])) AND (NOT D[1]))) OR D[2]) AND ((NOT ((D[4] AND (NOT D[3])) AND (NOT D[1]))) OR D[6])) AND ((NOT (((NOT D[4]) AND D[3]) AND (NOT D[1]))) OR D[7])) AND ((NOT ((D[4] AND D[3]) AND (NOT D[1]))) OR D[5])) AND ((NOT (((NOT D[4]) AND (NOT D[3])) AND D[1])) OR D[10])) AND ((NOT ((D[4] AND (NOT D[3])) AND D[1])) OR D[8])) AND ((NOT (((NOT D[4]) AND D[3]) AND D[1])) OR D[9])) AND ((NOT ((D[4] AND D[3]) AND D[1])) OR D[11]));
    OutReady := 1;
    CollectInput(RESET:=TRUE);
  END_IF;
END_PROGRAM

CONFIGURATION Config0
  RESOURCE Res0 ON PLC
    TASK task0(INTERVAL := T#20ms,PRIORITY := 0);
    PROGRAM instance0 WITH task0 : Boiler;
  END_RESOURCE
END_CONFIGURATION

(* ---- 3-MUX_dados-chirp-paint.st ---- *)
(*
This code implements a shuffled multiplexer with 3 control bits.
The control bits are: Data[9], Data[1], Data[3]
The input bits are: Data[2], Data[5], Data[10], Data[6], Data[7], Data[4], Data[8], Data[11]

The symbolic expression is:
(((((((~((~(D[9]) & ~(D[1])) & ~(D[3])) | D[2]) & (~((D[9] & ~(D[1])) & ~(D[3])) | D[5])) & (~((~(D[9]) & D[1]) & ~(D[3])) | D[10])) & (~((D[9] & D[1]) & ~(D[3])) | D[6])) & (~((~(D[9]) & ~(D[1])) & D[3]) | D[7])) & (~((D[9] & ~(D[1])) & D[3]) | D[4])) & (~((~(D[9]) & D[1]) & D[3]) | D[8])) & (~((D[9] & D[1]) & D[3]) | D[11])

*)

FUNCTION_BLOCK F_CollectInput
  VAR_IN_OUT
      Data : ARRAY[1..15] OF BOOL;
  END_VAR
  VAR_INPUT
      TICK  : BOOL := 0;
      IN1   : BOOL := 0;
      IN2   : BOOL := 0;
      IN3   : BOOL := 0;
      IN4   : BOOL := 0;
      IN5   : BOOL := 0;
      RESET : BOOL := FALSE;
  END_VAR
  VAR_OUTPUT
      Finished : BOOL;
  END_VAR
  VAR
      j    : USINT := 1;
      tock : BOOL  := 0;
  END_VAR
  IF NOT RESET AND tock = NOT TICK THEN
      Data[j]   := IN1;
      Data[j+1] := IN2;
      Data[j+2] := IN3;
      Data[j+3] := IN4;
      Data[j+4] := IN5;
      j := j + 5;
      tock := TICK;
  ELSE
      j := 1;
      tock := 0;
  END_IF;
  Finished := (j > 15);
END_FUNCTION_BLOCK

PROGRAM Boiler
  VAR
    Data  : ARRAY[1..15] OF BOOL;
    Ready : BOOL;
    CollectInput : F_CollectInput;
  END_VAR
  VAR
    TICK     AT %IX1.0 : BOOL;
    IN1      AT %IX0.3 : BOOL;
    IN2      AT %IX0.4 : BOOL;
    IN3      AT %IX0.5 : BOOL;
    IN4      AT %IX0.6 : BOOL;
    IN5      AT %IX0.7 : BOOL;
    OutReady AT %QX0.0 : BOOL := FALSE;
    FeedNext AT %QX0.1 : BOOL := FALSE;
    Out      AT %QX0.2 : BOOL;
  END_VAR
  CollectInput(TICK:=TICK, IN1:=IN1, IN2:=IN2, IN3:=IN3, IN4:=IN4, IN5:=IN5);
  Ready := CollectInput.Finished;
  FeedNext := 1;
  IF Ready THEN
    Out := (((((((((NOT (((NOT D[9]) AND (NOT D[1])) AND (NOT D[3]))) OR D[2]) AND ((NOT ((D[9] AND (NOT D[1])) AND (NOT D[3]))) OR D[5])) AND ((NOT (((NOT D[9]) AND D[1]) AND (NOT D[3]))) OR D[10])) AND ((NOT ((D[9] AND D[1]) AND (NOT D[3]))) OR D[6])) AND ((NOT (((NOT D[9]) AND (NOT D[1])) AND D[3])) OR D[7])) AND ((NOT ((D[9] AND (NOT D[1])) AND D[3])) OR D[4])) AND ((NOT (((NOT D[9]) AND D[1]) AND D[3])) OR D[8])) AND ((NOT ((D[9] AND D[1]) AND D[3])) OR D[11]));
    OutReady := 1;
    CollectInput(RESET:=TRUE);
  END_IF;
END_PROGRAM

CONFIGURATION Config0
  RESOURCE Res0 ON PLC
    TASK task0(INTERVAL := T#20ms,PRIORITY := 0);
    PROGRAM instance0 WITH task0 : Boiler;
  END_RESOURCE
END_CONFIGURATION

(* ---- 3-MUX_dewed-sorer-gales.st ---- *)
(*
This code implements a shuffled multiplexer with 3 control bits.
The control bits are: Data[2], Data[3], Data[1]
The input bits are: Data[4], Data[5], Data[7], Data[6], Data[9], Data[10], Data[8], Data[11]

The symbolic expression is:
(((((((~((~(D[2]) & ~(D[3])) & ~(D[1])) | D[4]) & (~((D[2] & ~(D[3])) & ~(D[1])) | D[5])) & (~((~(D[2]) & D[3]) & ~(D[1])) | D[7])) & (~((D[2] & D[3]) & ~(D[1])) | D[6])) & (~((~(D[2]) & ~(D[3])) & D[1]) | D[9])) & (~((D[2] & ~(D[3])) & D[1]) | D[10])) & (~((~(D[2]) & D[3]) & D[1]) | D[8])) & (~((D[2] & D[3]) & D[1]) | D[11])

*)

FUNCTION_BLOCK F_CollectInput
  VAR_IN_OUT
      Data : ARRAY[1..15] OF BOOL;
  END_VAR
  VAR_INPUT
      TICK  : BOOL := 0;
      IN1   : BOOL := 0;
      IN2   : BOOL := 0;
      IN3   : BOOL := 0;
      IN4   : BOOL := 0;
      IN5   : BOOL := 0;
      RESET : BOOL := FALSE;
  END_VAR
  VAR_OUTPUT
      Finished : BOOL;
  END_VAR
  VAR
      j    : USINT := 1;
      tock : BOOL  := 0;
  END_VAR
  IF NOT RESET AND tock = NOT TICK THEN
      Data[j]   := IN1;
      Data[j+1] := IN2;
      Data[j+2] := IN3;
      Data[j+3] := IN4;
      Data[j+4] := IN5;
      j := j + 5;
      tock := TICK;
  ELSE
      j := 1;
      tock := 0;
  END_IF;
  Finished := (j > 15);
END_FUNCTION_BLOCK

PROGRAM Boiler
  VAR
    Data  : ARRAY[1..15] OF BOOL;
    Ready : BOOL;
    CollectInput : F_CollectInput;
  END_VAR
  VAR
    TICK     AT %IX1.0 : BOOL;
    IN1      AT %IX0.3 : BOOL;
    IN2      AT %IX0.4 : BOOL;
    IN3      AT %IX0.5 : BOOL;
    IN4      AT %IX0.6 : BOOL;
    IN5      AT %IX0.7 : BOOL;
    OutReady AT %QX0.0 : BOOL := FALSE;
    FeedNext AT %QX0.1 : BOOL := FALSE;
    Out      AT %QX0.2 : BOOL;
  END_VAR
  CollectInput(TICK:=TICK, IN1:=IN1, IN2:=IN2, IN3:=IN3, IN4:=IN4, IN5:=IN5);
  Ready := CollectInput.Finished;
  FeedNext := 1;
  IF Ready THEN
    Out := (((((((((NOT (((NOT D[2]) AND (NOT D[3])) AND (NOT D[1]))) OR D[4]) AND ((NOT ((D[2] AND (NOT D[3])) AND (NOT D[1]))) OR D[5])) AND ((NOT (((NOT D[2]) AND D[3]) AND (NOT D[1]))) OR D[7])) AND ((NOT ((D[2] AND D[3]) AND (NOT D[1]))) OR D[6])) AND ((NOT (((NOT D[2]) AND (NOT D[3])) AND D[1])) OR D[9])) AND ((NOT ((D[2] AND (NOT D[3])) AND D[1])) OR D[10])) AND ((NOT (((NOT D[2]) AND D[3]) AND D[1])) OR D[8])) AND ((NOT ((D[2] AND D[3]) AND D[1])) OR D[11]));
    OutReady := 1;
    CollectInput(RESET:=TRUE);
  END_IF;
END_PROGRAM

CONFIGURATION Config0
  RESOURCE Res0 ON PLC
    TASK task0(INTERVAL := T#20ms,PRIORITY := 0);
    PROGRAM instance0 WITH task0 : Boiler;
  END_RESOURCE
END_CONFIGURATION

(* ---- 3-MUX_dopes-stump-meets.st ---- *)
(*
This code implements a shuffled multiplexer with 3 control bits.
The control bits are: Data[5], Data[2], Data[6]
The input bits are: Data[1], Data[8], Data[4], Data[9], Data[7], Data[10], Data[3], Data[11]

The symbolic expression is:
(((((((~((~(D[5]) & ~(D[2])) & ~(D[6])) | D[1]) & (~((D[5] & ~(D[2])) & ~(D[6])) | D[8])) & (~((~(D[5]) & D[2]) & ~(D[6])) | D[4])) & (~((D[5] & D[2]) & ~(D[6])) | D[9])) & (~((~(D[5]) & ~(D[2])) & D[6]) | D[7])) & (~((D[5] & ~(D[2])) & D[6]) | D[10])) & (~((~(D[5]) & D[2]) & D[6]) | D[3])) & (~((D[5] & D[2]) & D[6]) | D[11])

*)

FUNCTION_BLOCK F_CollectInput
  VAR_IN_OUT
      Data : ARRAY[1..15] OF BOOL;
  END_VAR
  VAR_INPUT
      TICK  : BOOL := 0;
      IN1   : BOOL := 0;
      IN2   : BOOL := 0;
      IN3   : BOOL := 0;
      IN4   : BOOL := 0;
      IN5   : BOOL := 0;
      RESET : BOOL := FALSE;
  END_VAR
  VAR_OUTPUT
      Finished : BOOL;
  END_VAR
  VAR
      j    : USINT := 1;
      tock : BOOL  := 0;
  END_VAR
  IF NOT RESET AND tock = NOT TICK THEN
      Data[j]   := IN1;
      Data[j+1] := IN2;
      Data[j+2] := IN3;
      Data[j+3] := IN4;
      Data[j+4] := IN5;
      j := j + 5;
      tock := TICK;
  ELSE
      j := 1;
      tock := 0;
  END_IF;
  Finished := (j > 15);
END_FUNCTION_BLOCK

PROGRAM Boiler
  VAR
    Data  : ARRAY[1..15] OF BOOL;
    Ready : BOOL;
    CollectInput : F_CollectInput;
  END_VAR
  VAR
    TICK     AT %IX1.0 : BOOL;
    IN1      AT %IX0.3 : BOOL;
    IN2      AT %IX0.4 : BOOL;
    IN3      AT %IX0.5 : BOOL;
    IN4      AT %IX0.6 : BOOL;
    IN5      AT %IX0.7 : BOOL;
    OutReady AT %QX0.0 : BOOL := FALSE;
    FeedNext AT %QX0.1 : BOOL := FALSE;
    Out      AT %QX0.2 : BOOL;
  END_VAR
  CollectInput(TICK:=TICK, IN1:=IN1, IN2:=IN2, IN3:=IN3, IN4:=IN4, IN5:=IN5);
  Ready := CollectInput.Finished;
  FeedNext := 1;
  IF Ready THEN
    Out := (((((((((NOT (((NOT D[5]) AND (NOT D[2])) AND (NOT D[6]))) OR D[1]) AND ((NOT ((D[5] AND (NOT D[2])) AND (NOT D[6]))) OR D[8])) AND ((NOT (((NOT D[5]) AND D[2]) AND (NOT D[6]))) OR D[4])) AND ((NOT ((D[5] AND D[2]) AND (NOT D[6]))) OR D[9])) AND ((NOT (((NOT D[5]) AND (NOT D[2])) AND D[6])) OR D[7])) AND ((NOT ((D[5] AND (NOT D[2])) AND D[6])) OR D[10])) AND ((NOT (((NOT D[5]) AND D[2]) AND D[6])) OR D[3])) AND ((NOT ((D[5] AND D[2]) AND D[6])) OR D[11]));
    OutReady := 1;
    CollectInput(RESET:=TRUE);
  END_IF;
END_PROGRAM

CONFIGURATION Config0
  RESOURCE Res0 ON PLC
    TASK task0(INTERVAL := T#20ms,PRIORITY := 0);
    PROGRAM instance0 WITH task0 : Boiler;
  END_RESOURCE
END_CONFIGURATION

(* ---- 3-MUX_drear-jiffs-guise.st ---- *)
(*
This code implements a shuffled multiplexer with 3 control bits.
The control bits are: Data[5], Data[2], Data[3]
The input bits are: Data[1], Data[6], Data[4], Data[8], Data[7], Data[10], Data[9], Data[11]

The symbolic expression is:
(((((((~((~(D[5]) & ~(D[2])) & ~(D[3])) | D[1]) & (~((D[5] & ~(D[2])) & ~(D[3])) | D[6])) & (~((~(D[5]) & D[2]) & ~(D[3])) | D[4])) & (~((D[5] & D[2]) & ~(D[3])) | D[8])) & (~((~(D[5]) & ~(D[2])) & D[3]) | D[7])) & (~((D[5] & ~(D[2])) & D[3]) | D[10])) & (~((~(D[5]) & D[2]) & D[3]) | D[9])) & (~((D[5] & D[2]) & D[3]) | D[11])

*)

FUNCTION_BLOCK F_CollectInput
  VAR_IN_OUT
      Data : ARRAY[1..15] OF BOOL;
  END_VAR
  VAR_INPUT
      TICK  : BOOL := 0;
      IN1   : BOOL := 0;
      IN2   : BOOL := 0;
      IN3   : BOOL := 0;
      IN4   : BOOL := 0;
      IN5   : BOOL := 0;
      RESET : BOOL := FALSE;
  END_VAR
  VAR_OUTPUT
      Finished : BOOL;
  END_VAR
  VAR
      j    : USINT := 1;
      tock : BOOL  := 0;
  END_VAR
  IF NOT RESET AND tock = NOT TICK THEN
      Data[j]   := IN1;
      Data[j+1] := IN2;
      Data[j+2] := IN3;
      Data[j+3] := IN4;
      Data[j+4] := IN5;
      j := j + 5;
      tock := TICK;
  ELSE
      j := 1;
      tock := 0;
  END_IF;
  Finished := (j > 15);
END_FUNCTION_BLOCK

PROGRAM Boiler
  VAR
    Data  : ARRAY[1..15] OF BOOL;
    Ready : BOOL;
    CollectInput : F_CollectInput;
  END_VAR
  VAR
    TICK     AT %IX1.0 : BOOL;
    IN1      AT %IX0.3 : BOOL;
    IN2      AT %IX0.4 : BOOL;
    IN3      AT %IX0.5 : BOOL;
    IN4      AT %IX0.6 : BOOL;
    IN5      AT %IX0.7 : BOOL;
    OutReady AT %QX0.0 : BOOL := FALSE;
    FeedNext AT %QX0.1 : BOOL := FALSE;
    Out      AT %QX0.2 : BOOL;
  END_VAR
  CollectInput(TICK:=TICK, IN1:=IN1, IN2:=IN2, IN3:=IN3, IN4:=IN4, IN5:=IN5);
  Ready := CollectInput.Finished;
  FeedNext := 1;
  IF Ready THEN
    Out := (((((((((NOT (((NOT D[5]) AND (NOT D[2])) AND (NOT D[3]))) OR D[1]) AND ((NOT ((D[5] AND (NOT D[2])) AND (NOT D[3]))) OR D[6])) AND ((NOT (((NOT D[5]) AND D[2]) AND (NOT D[3]))) OR D[4])) AND ((NOT ((D[5] AND D[2]) AND (NOT D[3]))) OR D[8])) AND ((NOT (((NOT D[5]) AND (NOT D[2])) AND D[3])) OR D[7])) AND ((NOT ((D[5] AND (NOT D[2])) AND D[3])) OR D[10])) AND ((NOT (((NOT D[5]) AND D[2]) AND D[3])) OR D[9])) AND ((NOT ((D[5] AND D[2]) AND D[3])) OR D[11]));
    OutReady := 1;
    CollectInput(RESET:=TRUE);
  END_IF;
END_PROGRAM

CONFIGURATION Config0
  RESOURCE Res0 ON PLC
    TASK task0(INTERVAL := T#20ms,PRIORITY := 0);
    PROGRAM instance0 WITH task0 : Boiler;
  END_RESOURCE
END_CONFIGURATION

(* ---- 3-MUX_dusky-quals-gales.st ---- *)
(*
This code implements a shuffled multiplexer with 3 control bits.
The control bits are: Data[3], Data[4], Data[5]
The input bits are: Data[6], Data[9], Data[1], Data[7], Data[2], Data[8], Data[10], Data[11]

The symbolic expression is:
(((((((~((~(D[3]) & ~(D[4])) & ~(D[5])) | D[6]) & (~((D[3] & ~(D[4])) & ~(D[5])) | D[9])) & (~((~(D[3]) & D[4]) & ~(D[5])) | D[1])) & (~((D[3] & D[4]) & ~(D[5])) | D[7])) & (~((~(D[3]) & ~(D[4])) & D[5]) | D[2])) & (~((D[3] & ~(D[4])) & D[5]) | D[8])) & (~((~(D[3]) & D[4]) & D[5]) | D[10])) & (~((D[3] & D[4]) & D[5]) | D[11])

*)

FUNCTION_BLOCK F_CollectInput
  VAR_IN_OUT
      Data : ARRAY[1..15] OF BOOL;
  END_VAR
  VAR_INPUT
      TICK  : BOOL := 0;
      IN1   : BOOL := 0;
      IN2   : BOOL := 0;
      IN3   : BOOL := 0;
      IN4   : BOOL := 0;
      IN5   : BOOL := 0;
      RESET : BOOL := FALSE;
  END_VAR
  VAR_OUTPUT
      Finished : BOOL;
  END_VAR
  VAR
      j    : USINT := 1;
      tock : BOOL  := 0;
  END_VAR
  IF NOT RESET AND tock = NOT TICK THEN
      Data[j]   := IN1;
      Data[j+1] := IN2;
      Data[j+2] := IN3;
      Data[j+3] := IN4;
      Data[j+4] := IN5;
      j := j + 5;
      tock := TICK;
  ELSE
      j := 1;
      tock := 0;
  END_IF;
  Finished := (j > 15);
END_FUNCTION_BLOCK

PROGRAM Boiler
  VAR
    Data  : ARRAY[1..15] OF BOOL;
    Ready : BOOL;
    CollectInput : F_CollectInput;
  END_VAR
  VAR
    TICK     AT %IX1.0 : BOOL;
    IN1      AT %IX0.3 : BOOL;
    IN2      AT %IX0.4 : BOOL;
    IN3      AT %IX0.5 : BOOL;
    IN4      AT %IX0.6 : BOOL;
    IN5      AT %IX0.7 : BOOL;
    OutReady AT %QX0.0 : BOOL := FALSE;
    FeedNext AT %QX0.1 : BOOL := FALSE;
    Out      AT %QX0.2 : BOOL;
  END_VAR
  CollectInput(TICK:=TICK, IN1:=IN1, IN2:=IN2, IN3:=IN3, IN4:=IN4, IN5:=IN5);
  Ready := CollectInput.Finished;
  FeedNext := 1;
  IF Ready THEN
    Out := (((((((((NOT (((NOT D[3]) AND (NOT D[4])) AND (NOT D[5]))) OR D[6]) AND ((NOT ((D[3] AND (NOT D[4])) AND (NOT D[5]))) OR D[9])) AND ((NOT (((NOT D[3]) AND D[4]) AND (NOT D[5]))) OR D[1])) AND ((NOT ((D[3] AND D[4]) AND (NOT D[5]))) OR D[7])) AND ((NOT (((NOT D[3]) AND (NOT D[4])) AND D[5])) OR D[2])) AND ((NOT ((D[3] AND (NOT D[4])) AND D[5])) OR D[8])) AND ((NOT (((NOT D[3]) AND D[4]) AND D[5])) OR D[10])) AND ((NOT ((D[3] AND D[4]) AND D[5])) OR D[11]));
    OutReady := 1;
    CollectInput(RESET:=TRUE);
  END_IF;
END_PROGRAM

CONFIGURATION Config0
  RESOURCE Res0 ON PLC
    TASK task0(INTERVAL := T#20ms,PRIORITY := 0);
    PROGRAM instance0 WITH task0 : Boiler;
  END_RESOURCE
END_CONFIGURATION

(* ---- 3-MUX_epsom-flies-chard.st ---- *)
(*
This code implements a shuffled multiplexer with 3 control bits.
The control bits are: Data[5], Data[2], Data[3]
The input bits are: Data[4], Data[1], Data[8], Data[7], Data[9], Data[6], Data[11], Data[10]

The symbolic expression is:
(((((((~((~(D[5]) & ~(D[2])) & ~(D[3])) | D[4]) & (~((D[5] & ~(D[2])) & ~(D[3])) | D[1])) & (~((~(D[5]) & D[2]) & ~(D[3])) | D[8])) & (~((D[5] & D[2]) & ~(D[3])) | D[7])) & (~((~(D[5]) & ~(D[2])) & D[3]) | D[9])) & (~((D[5] & ~(D[2])) & D[3]) | D[6])) & (~((~(D[5]) & D[2]) & D[3]) | D[11])) & (~((D[5] & D[2]) & D[3]) | D[10])

*)

FUNCTION_BLOCK F_CollectInput
  VAR_IN_OUT
      Data : ARRAY[1..15] OF BOOL;
  END_VAR
  VAR_INPUT
      TICK  : BOOL := 0;
      IN1   : BOOL := 0;
      IN2   : BOOL := 0;
      IN3   : BOOL := 0;
      IN4   : BOOL := 0;
      IN5   : BOOL := 0;
      RESET : BOOL := FALSE;
  END_VAR
  VAR_OUTPUT
      Finished : BOOL;
  END_VAR
  VAR
      j    : USINT := 1;
      tock : BOOL  := 0;
  END_VAR
  IF NOT RESET AND tock = NOT TICK THEN
      Data[j]   := IN1;
      Data[j+1] := IN2;
      Data[j+2] := IN3;
      Data[j+3] := IN4;
      Data[j+4] := IN5;
      j := j + 5;
      tock := TICK;
  ELSE
      j := 1;
      tock := 0;
  END_IF;
  Finished := (j > 15);
END_FUNCTION_BLOCK

PROGRAM Boiler
  VAR
    Data  : ARRAY[1..15] OF BOOL;
    Ready : BOOL;
    CollectInput : F_CollectInput;
  END_VAR
  VAR
    TICK     AT %IX1.0 : BOOL;
    IN1      AT %IX0.3 : BOOL;
    IN2      AT %IX0.4 : BOOL;
    IN3      AT %IX0.5 : BOOL;
    IN4      AT %IX0.6 : BOOL;
    IN5      AT %IX0.7 : BOOL;
    OutReady AT %QX0.0 : BOOL := FALSE;
    FeedNext AT %QX0.1 : BOOL := FALSE;
    Out      AT %QX0.2 : BOOL;
  END_VAR
  CollectInput(TICK:=TICK, IN1:=IN1, IN2:=IN2, IN3:=IN3, IN4:=IN4, IN5:=IN5);
  Ready := CollectInput.Finished;
  FeedNext := 1;
  IF Ready THEN
    Out := (((((((((NOT (((NOT D[5]) AND (NOT D[2])) AND (NOT D[3]))) OR D[4]) AND ((NOT ((D[5] AND (NOT D[2])) AND (NOT D[3]))) OR D[1])) AND ((NOT (((NOT D[5]) AND D[2]) AND (NOT D[3]))) OR D[8])) AND ((NOT ((D[5] AND D[2]) AND (NOT D[3]))) OR D[7])) AND ((NOT (((NOT D[5]) AND (NOT D[2])) AND D[3])) OR D[9])) AND ((NOT ((D[5] AND (NOT D[2])) AND D[3])) OR D[6])) AND ((NOT (((NOT D[5]) AND D[2]) AND D[3])) OR D[11])) AND ((NOT ((D[5] AND D[2]) AND D[3])) OR D[10]));
    OutReady := 1;
    CollectInput(RESET:=TRUE);
  END_IF;
END_PROGRAM

CONFIGURATION Config0
  RESOURCE Res0 ON PLC
    TASK task0(INTERVAL := T#20ms,PRIORITY := 0);
    PROGRAM instance0 WITH task0 : Boiler;
  END_RESOURCE
END_CONFIGURATION

(* ---- 3-MUX_erred-sprue-hodad.st ---- *)
(*
This code implements a shuffled multiplexer with 3 control bits.
The control bits are: Data[2], Data[3], Data[4]
The input bits are: Data[6], Data[1], Data[10], Data[5], Data[7], Data[9], Data[8], Data[11]

The symbolic expression is:
(((((((~((~(D[2]) & ~(D[3])) & ~(D[4])) | D[6]) & (~((D[2] & ~(D[3])) & ~(D[4])) | D[1])) & (~((~(D[2]) & D[3]) & ~(D[4])) | D[10])) & (~((D[2] & D[3]) & ~(D[4])) | D[5])) & (~((~(D[2]) & ~(D[3])) & D[4]) | D[7])) & (~((D[2] & ~(D[3])) & D[4]) | D[9])) & (~((~(D[2]) & D[3]) & D[4]) | D[8])) & (~((D[2] & D[3]) & D[4]) | D[11])

*)

FUNCTION_BLOCK F_CollectInput
  VAR_IN_OUT
      Data : ARRAY[1..15] OF BOOL;
  END_VAR
  VAR_INPUT
      TICK  : BOOL := 0;
      IN1   : BOOL := 0;
      IN2   : BOOL := 0;
      IN3   : BOOL := 0;
      IN4   : BOOL := 0;
      IN5   : BOOL := 0;
      RESET : BOOL := FALSE;
  END_VAR
  VAR_OUTPUT
      Finished : BOOL;
  END_VAR
  VAR
      j    : USINT := 1;
      tock : BOOL  := 0;
  END_VAR
  IF NOT RESET AND tock = NOT TICK THEN
      Data[j]   := IN1;
      Data[j+1] := IN2;
      Data[j+2] := IN3;
      Data[j+3] := IN4;
      Data[j+4] := IN5;
      j := j + 5;
      tock := TICK;
  ELSE
      j := 1;
      tock := 0;
  END_IF;
  Finished := (j > 15);
END_FUNCTION_BLOCK

PROGRAM Boiler
  VAR
    Data  : ARRAY[1..15] OF BOOL;
    Ready : BOOL;
    CollectInput : F_CollectInput;
  END_VAR
  VAR
    TICK     AT %IX1.0 : BOOL;
    IN1      AT %IX0.3 : BOOL;
    IN2      AT %IX0.4 : BOOL;
    IN3      AT %IX0.5 : BOOL;
    IN4      AT %IX0.6 : BOOL;
    IN5      AT %IX0.7 : BOOL;
    OutReady AT %QX0.0 : BOOL := FALSE;
    FeedNext AT %QX0.1 : BOOL := FALSE;
    Out      AT %QX0.2 : BOOL;
  END_VAR
  CollectInput(TICK:=TICK, IN1:=IN1, IN2:=IN2, IN3:=IN3, IN4:=IN4, IN5:=IN5);
  Ready := CollectInput.Finished;
  FeedNext := 1;
  IF Ready THEN
    Out := (((((((((NOT (((NOT D[2]) AND (NOT D[3])) AND (NOT D[4]))) OR D[6]) AND ((NOT ((D[2] AND (NOT D[3])) AND (NOT D[4]))) OR D[1])) AND ((NOT (((NOT D[2]) AND D[3]) AND (NOT D[4]))) OR D[10])) AND ((NOT ((D[2] AND D[3]) AND (NOT D[4]))) OR D[5])) AND ((NOT (((NOT D[2]) AND (NOT D[3])) AND D[4])) OR D[7])) AND ((NOT ((D[2] AND (NOT D[3])) AND D[4])) OR D[9])) AND ((NOT (((NOT D[2]) AND D[3]) AND D[4])) OR D[8])) AND ((NOT ((D[2] AND D[3]) AND D[4])) OR D[11]));
    OutReady := 1;
    CollectInput(RESET:=TRUE);
  END_IF;
END_PROGRAM

CONFIGURATION Config0
  RESOURCE Res0 ON PLC
    TASK task0(INTERVAL := T#20ms,PRIORITY := 0);
    PROGRAM instance0 WITH task0 : Boiler;
  END_RESOURCE
END_CONFIGURATION

(* ---- 3-MUX_etext-amuck-dined.st ---- *)
(*
This code implements a shuffled multiplexer with 3 control bits.
The control bits are: Data[4], Data[3], Data[2]
The input bits are: Data[5], Data[1], Data[7], Data[8], Data[6], Data[9], Data[10], Data[11]

The symbolic expression is:
(((((((~((~(D[4]) & ~(D[3])) & ~(D[2])) | D[5]) & (~((D[4] & ~(D[3])) & ~(D[2])) | D[1])) & (~((~(D[4]) & D[3]) & ~(D[2])) | D[7])) & (~((D[4] & D[3]) & ~(D[2])) | D[8])) & (~((~(D[4]) & ~(D[3])) & D[2]) | D[6])) & (~((D[4] & ~(D[3])) & D[2]) | D[9])) & (~((~(D[4]) & D[3]) & D[2]) | D[10])) & (~((D[4] & D[3]) & D[2]) | D[11])

*)

FUNCTION_BLOCK F_CollectInput
  VAR_IN_OUT
      Data : ARRAY[1..15] OF BOOL;
  END_VAR
  VAR_INPUT
      TICK  : BOOL := 0;
      IN1   : BOOL := 0;
      IN2   : BOOL := 0;
      IN3   : BOOL := 0;
      IN4   : BOOL := 0;
      IN5   : BOOL := 0;
      RESET : BOOL := FALSE;
  END_VAR
  VAR_OUTPUT
      Finished : BOOL;
  END_VAR
  VAR
      j    : USINT := 1;
      tock : BOOL  := 0;
  END_VAR
  IF NOT RESET AND tock = NOT TICK THEN
      Data[j]   := IN1;
      Data[j+1] := IN2;
      Data[j+2] := IN3;
      Data[j+3] := IN4;
      Data[j+4] := IN5;
      j := j + 5;
      tock := TICK;
  ELSE
      j := 1;
      tock := 0;
  END_IF;
  Finished := (j > 15);
END_FUNCTION_BLOCK

PROGRAM Boiler
  VAR
    Data  : ARRAY[1..15] OF BOOL;
    Ready : BOOL;
    CollectInput : F_CollectInput;
  END_VAR
  VAR
    TICK     AT %IX1.0 : BOOL;
    IN1      AT %IX0.3 : BOOL;
    IN2      AT %IX0.4 : BOOL;
    IN3      AT %IX0.5 : BOOL;
    IN4      AT %IX0.6 : BOOL;
    IN5      AT %IX0.7 : BOOL;
    OutReady AT %QX0.0 : BOOL := FALSE;
    FeedNext AT %QX0.1 : BOOL := FALSE;
    Out      AT %QX0.2 : BOOL;
  END_VAR
  CollectInput(TICK:=TICK, IN1:=IN1, IN2:=IN2, IN3:=IN3, IN4:=IN4, IN5:=IN5);
  Ready := CollectInput.Finished;
  FeedNext := 1;
  IF Ready THEN
    Out := (((((((((NOT (((NOT D[4]) AND (NOT D[3])) AND (NOT D[2]))) OR D[5]) AND ((NOT ((D[4] AND (NOT D[3])) AND (NOT D[2]))) OR D[1])) AND ((NOT (((NOT D[4]) AND D[3]) AND (NOT D[2]))) OR D[7])) AND ((NOT ((D[4] AND D[3]) AND (NOT D[2]))) OR D[8])) AND ((NOT (((NOT D[4]) AND (NOT D[3])) AND D[2])) OR D[6])) AND ((NOT ((D[4] AND (NOT D[3])) AND D[2])) OR D[9])) AND ((NOT (((NOT D[4]) AND D[3]) AND D[2])) OR D[10])) AND ((NOT ((D[4] AND D[3]) AND D[2])) OR D[11]));
    OutReady := 1;
    CollectInput(RESET:=TRUE);
  END_IF;
END_PROGRAM

CONFIGURATION Config0
  RESOURCE Res0 ON PLC
    TASK task0(INTERVAL := T#20ms,PRIORITY := 0);
    PROGRAM instance0 WITH task0 : Boiler;
  END_RESOURCE
END_CONFIGURATION

(* ---- 3-MUX_filch-foods-lipid.st ---- *)
(*
This code implements a shuffled multiplexer with 3 control bits.
The control bits are: Data[3], Data[2], Data[1]
The input bits are: Data[4], Data[7], Data[5], Data[8], Data[6], Data[9], Data[10], Data[11]

The symbolic expression is:
(((((((~((~(D[3]) & ~(D[2])) & ~(D[1])) | D[4]) & (~((D[3] & ~(D[2])) & ~(D[1])) | D[7])) & (~((~(D[3]) & D[2]) & ~(D[1])) | D[5])) & (~((D[3] & D[2]) & ~(D[1])) | D[8])) & (~((~(D[3]) & ~(D[2])) & D[1]) | D[6])) & (~((D[3] & ~(D[2])) & D[1]) | D[9])) & (~((~(D[3]) & D[2]) & D[1]) | D[10])) & (~((D[3] & D[2]) & D[1]) | D[11])

*)

FUNCTION_BLOCK F_CollectInput
  VAR_IN_OUT
      Data : ARRAY[1..15] OF BOOL;
  END_VAR
  VAR_INPUT
      TICK  : BOOL := 0;
      IN1   : BOOL := 0;
      IN2   : BOOL := 0;
      IN3   : BOOL := 0;
      IN4   : BOOL := 0;
      IN5   : BOOL := 0;
      RESET : BOOL := FALSE;
  END_VAR
  VAR_OUTPUT
      Finished : BOOL;
  END_VAR
  VAR
      j    : USINT := 1;
      tock : BOOL  := 0;
  END_VAR
  IF NOT RESET AND tock = NOT TICK THEN
      Data[j]   := IN1;
      Data[j+1] := IN2;
      Data[j+2] := IN3;
      Data[j+3] := IN4;
      Data[j+4] := IN5;
      j := j + 5;
      tock := TICK;
  ELSE
      j := 1;
      tock := 0;
  END_IF;
  Finished := (j > 15);
END_FUNCTION_BLOCK

PROGRAM Boiler
  VAR
    Data  : ARRAY[1..15] OF BOOL;
    Ready : BOOL;
    CollectInput : F_CollectInput;
  END_VAR
  VAR
    TICK     AT %IX1.0 : BOOL;
    IN1      AT %IX0.3 : BOOL;
    IN2      AT %IX0.4 : BOOL;
    IN3      AT %IX0.5 : BOOL;
    IN4      AT %IX0.6 : BOOL;
    IN5      AT %IX0.7 : BOOL;
    OutReady AT %QX0.0 : BOOL := FALSE;
    FeedNext AT %QX0.1 : BOOL := FALSE;
    Out      AT %QX0.2 : BOOL;
  END_VAR
  CollectInput(TICK:=TICK, IN1:=IN1, IN2:=IN2, IN3:=IN3, IN4:=IN4, IN5:=IN5);
  Ready := CollectInput.Finished;
  FeedNext := 1;
  IF Ready THEN
    Out := (((((((((NOT (((NOT D[3]) AND (NOT D[2])) AND (NOT D[1]))) OR D[4]) AND ((NOT ((D[3] AND (NOT D[2])) AND (NOT D[1]))) OR D[7])) AND ((NOT (((NOT D[3]) AND D[2]) AND (NOT D[1]))) OR D[5])) AND ((NOT ((D[3] AND D[2]) AND (NOT D[1]))) OR D[8])) AND ((NOT (((NOT D[3]) AND (NOT D[2])) AND D[1])) OR D[6])) AND ((NOT ((D[3] AND (NOT D[2])) AND D[1])) OR D[9])) AND ((NOT (((NOT D[3]) AND D[2]) AND D[1])) OR D[10])) AND ((NOT ((D[3] AND D[2]) AND D[1])) OR D[11]));
    OutReady := 1;
    CollectInput(RESET:=TRUE);
  END_IF;
END_PROGRAM

CONFIGURATION Config0
  RESOURCE Res0 ON PLC
    TASK task0(INTERVAL := T#20ms,PRIORITY := 0);
    PROGRAM instance0 WITH task0 : Boiler;
  END_RESOURCE
END_CONFIGURATION

(* ---- 3-MUX_filth-genet-crack.st ---- *)
(*
This code implements a shuffled multiplexer with 3 control bits.
The control bits are: Data[2], Data[3], Data[1]
The input bits are: Data[4], Data[5], Data[6], Data[7], Data[9], Data[10], Data[8], Data[11]

The symbolic expression is:
(((((((~((~(D[2]) & ~(D[3])) & ~(D[1])) | D[4]) & (~((D[2] & ~(D[3])) & ~(D[1])) | D[5])) & (~((~(D[2]) & D[3]) & ~(D[1])) | D[6])) & (~((D[2] & D[3]) & ~(D[1])) | D[7])) & (~((~(D[2]) & ~(D[3])) & D[1]) | D[9])) & (~((D[2] & ~(D[3])) & D[1]) | D[10])) & (~((~(D[2]) & D[3]) & D[1]) | D[8])) & (~((D[2] & D[3]) & D[1]) | D[11])

*)

FUNCTION_BLOCK F_CollectInput
  VAR_IN_OUT
      Data : ARRAY[1..15] OF BOOL;
  END_VAR
  VAR_INPUT
      TICK  : BOOL := 0;
      IN1   : BOOL := 0;
      IN2   : BOOL := 0;
      IN3   : BOOL := 0;
      IN4   : BOOL := 0;
      IN5   : BOOL := 0;
      RESET : BOOL := FALSE;
  END_VAR
  VAR_OUTPUT
      Finished : BOOL;
  END_VAR
  VAR
      j    : USINT := 1;
      tock : BOOL  := 0;
  END_VAR
  IF NOT RESET AND tock = NOT TICK THEN
      Data[j]   := IN1;
      Data[j+1] := IN2;
      Data[j+2] := IN3;
      Data[j+3] := IN4;
      Data[j+4] := IN5;
      j := j + 5;
      tock := TICK;
  ELSE
      j := 1;
      tock := 0;
  END_IF;
  Finished := (j > 15);
END_FUNCTION_BLOCK

PROGRAM Boiler
  VAR
    Data  : ARRAY[1..15] OF BOOL;
    Ready : BOOL;
    CollectInput : F_CollectInput;
  END_VAR
  VAR
    TICK     AT %IX1.0 : BOOL;
    IN1      AT %IX0.3 : BOOL;
    IN2      AT %IX0.4 : BOOL;
    IN3      AT %IX0.5 : BOOL;
    IN4      AT %IX0.6 : BOOL;
    IN5      AT %IX0.7 : BOOL;
    OutReady AT %QX0.0 : BOOL := FALSE;
    FeedNext AT %QX0.1 : BOOL := FALSE;
    Out      AT %QX0.2 : BOOL;
  END_VAR
  CollectInput(TICK:=TICK, IN1:=IN1, IN2:=IN2, IN3:=IN3, IN4:=IN4, IN5:=IN5);
  Ready := CollectInput.Finished;
  FeedNext := 1;
  IF Ready THEN
    Out := (((((((((NOT (((NOT D[2]) AND (NOT D[3])) AND (NOT D[1]))) OR D[4]) AND ((NOT ((D[2] AND (NOT D[3])) AND (NOT D[1]))) OR D[5])) AND ((NOT (((NOT D[2]) AND D[3]) AND (NOT D[1]))) OR D[6])) AND ((NOT ((D[2] AND D[3]) AND (NOT D[1]))) OR D[7])) AND ((NOT (((NOT D[2]) AND (NOT D[3])) AND D[1])) OR D[9])) AND ((NOT ((D[2] AND (NOT D[3])) AND D[1])) OR D[10])) AND ((NOT (((NOT D[2]) AND D[3]) AND D[1])) OR D[8])) AND ((NOT ((D[2] AND D[3]) AND D[1])) OR D[11]));
    OutReady := 1;
    CollectInput(RESET:=TRUE);
  END_IF;
END_PROGRAM

CONFIGURATION Config0
  RESOURCE Res0 ON PLC
    TASK task0(INTERVAL := T#20ms,PRIORITY := 0);
    PROGRAM instance0 WITH task0 : Boiler;
  END_RESOURCE
END_CONFIGURATION

(* ---- 3-MUX_finds-mango-atoll.st ---- *)
(*
This code implements a shuffled multiplexer with 3 control bits.
The control bits are: Data[4], Data[1], Data[3]
The input bits are: Data[6], Data[2], Data[5], Data[7], Data[11], Data[8], Data[9], Data[10]

The symbolic expression is:
(((((((~((~(D[4]) & ~(D[1])) & ~(D[3])) | D[6]) & (~((D[4] & ~(D[1])) & ~(D[3])) | D[2])) & (~((~(D[4]) & D[1]) & ~(D[3])) | D[5])) & (~((D[4] & D[1]) & ~(D[3])) | D[7])) & (~((~(D[4]) & ~(D[1])) & D[3]) | D[11])) & (~((D[4] & ~(D[1])) & D[3]) | D[8])) & (~((~(D[4]) & D[1]) & D[3]) | D[9])) & (~((D[4] & D[1]) & D[3]) | D[10])

*)

FUNCTION_BLOCK F_CollectInput
  VAR_IN_OUT
      Data : ARRAY[1..15] OF BOOL;
  END_VAR
  VAR_INPUT
      TICK  : BOOL := 0;
      IN1   : BOOL := 0;
      IN2   : BOOL := 0;
      IN3   : BOOL := 0;
      IN4   : BOOL := 0;
      IN5   : BOOL := 0;
      RESET : BOOL := FALSE;
  END_VAR
  VAR_OUTPUT
      Finished : BOOL;
  END_VAR
  VAR
      j    : USINT := 1;
      tock : BOOL  := 0;
  END_VAR
  IF NOT RESET AND tock = NOT TICK THEN
      Data[j]   := IN1;
      Data[j+1] := IN2;
      Data[j+2] := IN3;
      Data[j+3] := IN4;
      Data[j+4] := IN5;
      j := j + 5;
      tock := TICK;
  ELSE
      j := 1;
      tock := 0;
  END_IF;
  Finished := (j > 15);
END_FUNCTION_BLOCK

PROGRAM Boiler
  VAR
    Data  : ARRAY[1..15] OF BOOL;
    Ready : BOOL;
    CollectInput : F_CollectInput;
  END_VAR
  VAR
    TICK     AT %IX1.0 : BOOL;
    IN1      AT %IX0.3 : BOOL;
    IN2      AT %IX0.4 : BOOL;
    IN3      AT %IX0.5 : BOOL;
    IN4      AT %IX0.6 : BOOL;
    IN5      AT %IX0.7 : BOOL;
    OutReady AT %QX0.0 : BOOL := FALSE;
    FeedNext AT %QX0.1 : BOOL := FALSE;
    Out      AT %QX0.2 : BOOL;
  END_VAR
  CollectInput(TICK:=TICK, IN1:=IN1, IN2:=IN2, IN3:=IN3, IN4:=IN4, IN5:=IN5);
  Ready := CollectInput.Finished;
  FeedNext := 1;
  IF Ready THEN
    Out := (((((((((NOT (((NOT D[4]) AND (NOT D[1])) AND (NOT D[3]))) OR D[6]) AND ((NOT ((D[4] AND (NOT D[1])) AND (NOT D[3]))) OR D[2])) AND ((NOT (((NOT D[4]) AND D[1]) AND (NOT D[3]))) OR D[5])) AND ((NOT ((D[4] AND D[1]) AND (NOT D[3]))) OR D[7])) AND ((NOT (((NOT D[4]) AND (NOT D[1])) AND D[3])) OR D[11])) AND ((NOT ((D[4] AND (NOT D[1])) AND D[3])) OR D[8])) AND ((NOT (((NOT D[4]) AND D[1]) AND D[3])) OR D[9])) AND ((NOT ((D[4] AND D[1]) AND D[3])) OR D[10]));
    OutReady := 1;
    CollectInput(RESET:=TRUE);
  END_IF;
END_PROGRAM

CONFIGURATION Config0
  RESOURCE Res0 ON PLC
    TASK task0(INTERVAL := T#20ms,PRIORITY := 0);
    PROGRAM instance0 WITH task0 : Boiler;
  END_RESOURCE
END_CONFIGURATION
